(* Q: 고르기 → 응답 필터 → 제한 (지령원 Q 제한 + 정격 + 제한 모듈 Q). 다른 경로 몫을 합쳐 제한 (Auto만) *)
stQRng := F_RangeOpen();
IF _stApply.bSrcLimit THEN
	stQRng := _stQSrcLim;		// 지령원 Q 제한 (P와 같음: Manual은 정책 bSrcLimit). 접속점 기준 → 설비 기준 (보정만큼 옮김)
	IF stQRng.nMaxModule <> 0 THEN stQRng.fMax := stQRng.fMax + fQComp; END_IF
	IF stQRng.nMinModule <> 0 THEN stQRng.fMin := stQRng.fMin + fQComp; END_IF
END_IF
IF _stApply.bRating THEN
	stQRng := F_RangeAnd(stQRng, _stEnv.stQ);
END_IF
FOR i := 1 TO GVL_PARAM.LIMIT_COUNT DO
	// Q도 P와 같은 규칙: 설비 기준 모듈은 bDevLimit, 접속점 기준 모듈은 M_PccLimitOn (Manual은 bPccLimit + 모듈 bManual)
	// Q 범위는 설비 기준(접속점 + 보정)이므로 접속점 기준 모듈 값은 보정만큼 옮겨 겹침 (P는 보정 앞 단계에서 자름)
	IF M_DevLimitOn(i) THEN
		stQRng := F_RangeAdd(stQRng, _astLim[i].stQ, _anLimModule[i]);
	ELSIF M_PccLimitOn(i) THEN
		stQLim		:= _astLim[i].stQ;
		stQLim.fMax	:= stQLim.fMax + fQComp;
		stQLim.fMin	:= stQLim.fMin + fQComp;
		stQRng := F_RangeAdd(stQRng, stQLim, _anLimModule[i]);
	END_IF
END_FOR
stDiag.stQRng		:= stQRng;
stDiag.bQGroupCmd	:= _stGrpQ.bActive;
stDiag.bQUnitCmd	:= _bUnitQCmd;
tTau := T#0S;
IF _stApply.bRamp THEN
	tTau := _tQFilter;
END_IF
// 목표 = 그룹 지령 (필터 후 + 보정). 없으면 유닛 지령 합 + 다른 경로 몫 (필터는 그 값을 따라가게만 둠)
IF _stGrpQ.bActive THEN
	_afbQFilter[i_nGroup](i_fIn := _stGrpQ.fValue, i_tTau := tTau);
	stDiag.stQ := F_RangeClamp(_afbQFilter[i_nGroup].q_fOut + fQComp, stQRng);
ELSE
	_afbQFilter[i_nGroup](i_fIn := _fUnitQSum + _fOtherQ - fQComp, i_tTau := tTau);
	stDiag.stQ := F_RangeClamp(_fUnitQSum + _fOtherQ, stQRng);
END_IF
M_ShapePath := stDiag;
END_METHOD

METHOD PRIVATE M_PccLimitOn : BOOL		// 이번 경로에 접속점 기준 모듈 i를 적용하는가
VAR_INPUT
	i_nLimit	: UINT;
END_VAR
M_PccLimitOn := _abLimOn[i_nLimit] AND _aeBasis[i_nLimit] = E_LimitBasis.Pcc
				AND (NOT i_bManual OR (_stApply.bPccLimit AND _abPccManual[i_nLimit]));
END_METHOD

METHOD PRIVATE M_DevLimitOn : BOOL		// 이번 경로에 설비 기준 모듈 i를 적용하는가 (Manual은 정책 bDevLimit)
VAR_INPUT
	i_nLimit	: UINT;
END_VAR
M_DevLimitOn := _stApply.bDevLimit AND _abLimOn[i_nLimit] AND _aeBasis[i_nLimit] = E_LimitBasis.Device;
END_METHOD

METHOD PRIVATE M_TraceSet		// 추적표에 한 줄 추가
VAR_INPUT
	i_eStep		: E_TraceStep;
	i_fValue	: REAL;
	i_nModule	: UINT;
	i_bCut		: BOOL;
END_VAR
IF _stTrace.nCount < GVL_PARAM.TRACE_STEP_MAX - 2 THEN		// 끝 두 줄(분배 후·쓴 값)은 FB_OutputDiag 몫
	_stTrace.nCount := _stTrace.nCount + 1;
	_stTrace.astStep[_stTrace.nCount].eStep		:= i_eStep;
	_stTrace.astStep[_stTrace.nCount].fValue	:= i_fValue;
	_stTrace.astStep[_stTrace.nCount].bCut		:= i_bCut;
	_stTrace.astStep[_stTrace.nCount].nModule	:= i_nModule;
	_stTrace.astStep[_stTrace.nCount].nReason	:= 0;
END_IF
END_METHOD

METHOD PRIVATE M_TraceClamp : REAL		// 범위 하나로 자르고 추적표에 한 줄. 자른 값을 돌려줌
VAR_INPUT
	i_eStep		: E_TraceStep;
	i_fIn		: REAL;
	i_stRange	: ST_Range;
END_VAR
VAR
	stClamp		: ST_Clamp;
END_VAR
stClamp := F_RangeClamp(i_fIn, i_stRange);
M_TraceSet(i_eStep, stClamp.fOut, stClamp.nModule, stClamp.bClamped);
IF _stTrace.nCount >= 1 THEN
	_stTrace.astStep[_stTrace.nCount].nReason := stClamp.nReason;
END_IF
M_TraceClamp := stClamp.fOut;
END_METHOD

END_FUNCTION_BLOCK

// ---- 10_Core/02_Util/FB_Lpf.TcPOU
FUNCTION_BLOCK FB_Lpf		// 1차 지연 필터
VAR_INPUT
	i_fIn			: REAL;
	i_tTau			: TIME;		// 시정수. T#0S면 필터 없이 통과
	i_bSync			: BOOL;		// 내부 값을 i_fSyncValue로 맞춤
	i_fSyncValue	: REAL;
END_VAR
VAR_OUTPUT
	q_fOut			: REAL;
END_VAR
VAR
	_fState			: REAL;
END_VAR
VAR_TEMP
	fDt				: REAL;		// s
	fTau			: REAL;		// s
END_VAR

fDt		:= F_CycleSec();
fTau	:= TIME_TO_REAL(i_tTau) / 1000.0;

IF i_bSync THEN
	_fState := i_fSyncValue;
ELSIF fTau <= 0 THEN
	_fState := i_fIn;
ELSE
	_fState := _fState + (fDt / (fTau + fDt)) * (i_fIn - _fState);
END_IF

q_fOut := _fState;

END_FUNCTION_BLOCK

// ---- 10_Core/02_Util/F_CycleSec.TcPOU
FUNCTION F_CycleSec : REAL		// 지금 태스크의 주기 (s)
VAR
	nTask		: DINT;
END_VAR

nTask := GETCURTASKINDEXEX();
F_CycleSec := UDINT_TO_REAL(TwinCAT_SystemInfoVarList._TaskInfo[nTask].CycleTime) * 1.0E-7;	// 100 ns 단위

END_FUNCTION

// ---- 10_Core/02_Util/F_RampStep.TcPOU
FUNCTION F_RampStep : REAL		// 기준값에서 한 스캔 동안 갈 수 있는 만큼만 목표 쪽으로
VAR_INPUT
	i_fTarget	: REAL;
	i_fRef		: REAL;			// 기준 (지난 스캔 최종 출력)
	i_fUpRate	: REAL;			// |값|이 커지는 쪽 (단위/s). 0 = 램프 없음
	i_fDnRate	: REAL;			// |값|이 작아지는 쪽 (단위/s). 0 = 램프 없음
END_VAR
VAR
	fRate		: REAL;
	fStep		: REAL;
END_VAR

IF ABS(i_fTarget) > ABS(i_fRef) AND i_fTarget * i_fRef >= 0 THEN
	fRate := i_fUpRate;
ELSE
	fRate := i_fDnRate;
END_IF

IF fRate <= 0 THEN
	F_RampStep := i_fTarget;
ELSE
	fStep		:= fRate * F_CycleSec();
	F_RampStep	:= i_fRef + LIMIT(-fStep, i_fTarget - i_fRef, fStep);
END_IF

END_FUNCTION

// ---- 10_Core/40_Arbitration/F_RangeClamp.TcPOU
FUNCTION F_RangeClamp : ST_Clamp		// 값을 범위 안으로. 상·하한이 겹치면 상한이 이김
VAR_INPUT
	i_fIn		: REAL;
	i_stRange	: ST_Range;
END_VAR

F_RangeClamp.fIn	:= i_fIn;
F_RangeClamp.fOut	:= i_fIn;
IF F_RangeClamp.fOut < i_stRange.fMin THEN
	F_RangeClamp.fOut		:= i_stRange.fMin;
	F_RangeClamp.bClamped	:= TRUE;
	F_RangeClamp.nModule	:= i_stRange.nMinModule;
	F_RangeClamp.nReason	:= i_stRange.nMinReason;
END_IF
IF F_RangeClamp.fOut > i_stRange.fMax THEN
	F_RangeClamp.fOut		:= i_stRange.fMax;
	F_RangeClamp.bClamped	:= TRUE;
	F_RangeClamp.nModule	:= i_stRange.nMaxModule;
	F_RangeClamp.nReason	:= i_stRange.nMaxReason;
END_IF

END_FUNCTION

// ---- 10_Core/50_Distribution/FB_Distributor.TcPOU
FUNCTION_BLOCK FB_Distributor		// 유닛에 나눔: 경로마다(Manual → Auto) 유닛 지령 → 그룹 몫 → 유닛 지령 축소, 그다음 배터리 그룹(방향·순 한도) → 피상전력
// Auto·Manual이 같은 순서 (M_DistPath). 그룹 지령이 없으면 그룹 몫은 0 (지령 없는 유닛은 0). 유닛 지령은 성형 결과(제한)에 걸릴 때만 줄임
// Manual 정책에서 정격·BMS 한도를 끈 Manual 유닛은 그 한도를 안 씀 (bRating을 끄면 유닛 제한 모듈만 씀)
// 유닛·버스 한도는 FB_EquipmentLimits 결과. 버스 한도는 나누는 동안 남은 한도로 보고(넘친 몫은 다른 유닛에 재분배), 끝에 한 번 더 확인
// 그룹 몫을 나누는 무게는 분배 정책(그룹마다 I_DistPolicy, 비우면 코어 기본 FB_DistStd = eDistBasis). 음수·이상값 무게는 0
VAR_IN_OUT
	iq_aipDistPolicy	: ARRAY[1..GVL_PARAM.GROUP_COUNT] OF I_DistPolicy;	// 그룹별 분배 정책 (GVL_SITE.g_aipDistPolicy)
END_VAR
VAR_IN_OUT CONSTANT
	(* Auto 경로 (fbAutoShape·fbAutoGate) *)
	iq_afAutoGrpP		: ARRAY[1..GVL_PARAM.GROUP_COUNT] OF REAL;
	iq_afAutoGrpQ		: ARRAY[1..GVL_PARAM.GROUP_COUNT] OF REAL;
	iq_afAutoUnitP		: ARRAY[1..GVL_PARAM.UNIT_COUNT] OF REAL;
	iq_afAutoUnitQ		: ARRAY[1..GVL_PARAM.UNIT_COUNT] OF REAL;
	iq_astAutoUnitP		: ARRAY[1..GVL_PARAM.UNIT_COUNT] OF ST_Pick;		// 유닛별 값이 있는지
	iq_astAutoUnitQ		: ARRAY[1..GVL_PARAM.UNIT_COUNT] OF ST_Pick;
	iq_abAutoGrpPCmd	: ARRAY[1..GVL_PARAM.GROUP_COUNT] OF BOOL;		// Auto 그룹 P 지령 있음 (fbAutoShape.q_abGrpPCmd)
	iq_abAutoGrpQCmd	: ARRAY[1..GVL_PARAM.GROUP_COUNT] OF BOOL;
	(* Manual 경로 (fbManualShape·fbManualGate) *)
	iq_afManualGrpP		: ARRAY[1..GVL_PARAM.GROUP_COUNT] OF REAL;
	iq_afManualGrpQ		: ARRAY[1..GVL_PARAM.GROUP_COUNT] OF REAL;
	iq_afManualUnitP	: ARRAY[1..GVL_PARAM.UNIT_COUNT] OF REAL;
	iq_afManualUnitQ	: ARRAY[1..GVL_PARAM.UNIT_COUNT] OF REAL;
	iq_astManualUnitP	: ARRAY[1..GVL_PARAM.UNIT_COUNT] OF ST_Pick;
	iq_astManualUnitQ	: ARRAY[1..GVL_PARAM.UNIT_COUNT] OF ST_Pick;
	iq_abManualGrpPCmd	: ARRAY[1..GVL_PARAM.GROUP_COUNT] OF BOOL;		// Manual 그룹 P 지령 있음 (fbManualShape.q_abGrpPCmd)
	iq_abManualGrpQCmd	: ARRAY[1..GVL_PARAM.GROUP_COUNT] OF BOOL;
	iq_astManualPolicy	: ARRAY[1..GVL_PARAM.GROUP_COUNT] OF ST_ManualPolicy;
	(* 공통 *)
	iq_abOutputReady	: ARRAY[1..GVL_PARAM.UNIT_COUNT] OF BOOL;	// 유닛 출력 가능 = 분배 대상 (FB_OutputReady)
	iq_aeNotReadyBy	: ARRAY[1..GVL_PARAM.UNIT_COUNT] OF E_UnitLimitBy;	// 못 내는 이유
	iq_aeOpMode		: ARRAY[1..GVL_PARAM.UNIT_COUNT] OF E_OpMode;
	iq_astUnitEnv	: ARRAY[1..GVL_PARAM.UNIT_COUNT] OF ST_UnitEnvelope;	// 유닛 한도 (FB_EquipmentLimits)
	iq_astBatEnv	: ARRAY[1..GVL_PARAM.BAT_COUNT] OF ST_BatEnvelope;	// 버스 한도 (FB_EquipmentLimits)
	iq_astUnitCfg	: ARRAY[1..GVL_PARAM.UNIT_COUNT] OF ST_UnitCfg;
	iq_astBatGroup	: ARRAY[1..GVL_PARAM.BAT_COUNT] OF ST_BatGroupState;
	iq_astGroupSet	: ARRAY[1..GVL_PARAM.GROUP_COUNT] OF ST_GroupSet;
END_VAR
VAR_OUTPUT
	q_astUnitSet	: ARRAY[1..GVL_PARAM.UNIT_COUNT] OF ST_PQ;		// 유닛 최종 지령
	q_astUnitDiag	: ARRAY[1..GVL_PARAM.UNIT_COUNT] OF ST_UnitDiag;
	q_astDistDiag	: ARRAY[1..GVL_PARAM.GROUP_COUNT] OF ST_DistDiag;
	q_astBatDiag	: ARRAY[1..GVL_PARAM.BAT_COUNT] OF ST_BatDistDiag;
	q_abUnitLimited	: ARRAY[1..GVL_PARAM.UNIT_COUNT] OF BOOL;		// 유닛 지령이 요청보다 줄었거나 0으로 묶임 (P 또는 Q). 제어용: Manual 재전송 판단 (FB_Dispatcher)
	q_abManualLimitOff: ARRAY[1..GVL_PARAM.GROUP_COUNT] OF BOOL;		// Manual 정책에서 정격·BMS 한도 중 하나라도 꺼짐 (HMI 표시용)
END_VAR
VAR
	(* 유닛 사본·작업값 (메서드에서 씀) *)
	_anGroup		: ARRAY[1..GVL_PARAM.UNIT_COUNT] OF UINT;
	_anBat			: ARRAY[1..GVL_PARAM.UNIT_COUNT] OF UINT;
	_abInDist		: ARRAY[1..GVL_PARAM.UNIT_COUNT] OF BOOL;		// 출력 가능 (FB_OutputReady)
	_abManual		: ARRAY[1..GVL_PARAM.UNIT_COUNT] OF BOOL;
	_abPFix			: ARRAY[1..GVL_PARAM.UNIT_COUNT] OF BOOL;		// 자기 경로에 유닛별 P 값 있음
	_abQFix			: ARRAY[1..GVL_PARAM.UNIT_COUNT] OF BOOL;
	_afPUnitReq		: ARRAY[1..GVL_PARAM.UNIT_COUNT] OF REAL;		// 자기 경로 유닛별 값 (성형 후)
	_afQUnitReq		: ARRAY[1..GVL_PARAM.UNIT_COUNT] OF REAL;
	_abNoRating		: ARRAY[1..GVL_PARAM.UNIT_COUNT] OF BOOL;		// Manual 정책: 정격·Derate·피상전력 안 씀
	_abNoBatLimit	: ARRAY[1..GVL_PARAM.UNIT_COUNT] OF BOOL;		// Manual 정책: BMS 충방전 한도 안 씀
	_astUnitEnv	: ARRAY[1..GVL_PARAM.UNIT_COUNT] OF ST_UnitEnvelope;	// 유닛 한도 사본 (메서드에서 씀)
	_astBatEnv	: ARRAY[1..GVL_PARAM.BAT_COUNT] OF ST_BatEnvelope;	// 버스 한도 사본
	_afBusDisLeft	: ARRAY[1..GVL_PARAM.BAT_COUNT] OF REAL;	// 버스 방전 쪽 남은 한도 (양수, 나누는 동안 줄어듦. 여러 그룹이 같은 버스를 써도 한 번만 씀)
	_afBusChgLeft	: ARRAY[1..GVL_PARAM.BAT_COUNT] OF REAL;	// 버스 충전 쪽 남은 한도 (양수)
	_anPModule	: ARRAY[1..GVL_PARAM.UNIT_COUNT] OF UINT;	// P를 줄인 모듈 (유닛 제한·버스 제한 모듈. 0 = 코어)
	_afPMax			: ARRAY[1..GVL_PARAM.UNIT_COUNT] OF REAL;
	_afPMin			: ARRAY[1..GVL_PARAM.UNIT_COUNT] OF REAL;
	_afQMax			: ARRAY[1..GVL_PARAM.UNIT_COUNT] OF REAL;
	_afQMin			: ARRAY[1..GVL_PARAM.UNIT_COUNT] OF REAL;
	_afPRated		: ARRAY[1..GVL_PARAM.UNIT_COUNT] OF REAL;
	_afQRated		: ARRAY[1..GVL_PARAM.UNIT_COUNT] OF REAL;
	_afSoc			: ARRAY[1..GVL_PARAM.UNIT_COUNT] OF REAL;		// 연결 배터리 그룹 SOC (%). 모르면 -1
	_afPWork		: ARRAY[1..GVL_PARAM.UNIT_COUNT] OF REAL;
	_afQWork		: ARRAY[1..GVL_PARAM.UNIT_COUNT] OF REAL;
	_aePBy			: ARRAY[1..GVL_PARAM.UNIT_COUNT] OF E_UnitLimitBy;
	_aeQBy			: ARRAY[1..GVL_PARAM.UNIT_COUNT] OF E_UnitLimitBy;
	_afPWeight		: ARRAY[1..GVL_PARAM.UNIT_COUNT] OF REAL;		// P 몫을 나눌 때 쓴 무게 (진단)
	_abBatNoChg		: ARRAY[1..GVL_PARAM.UNIT_COUNT] OF BOOL;		// 연결 배터리 버스 충전 한도 0 → 충전 몫 안 줌
	_abBatNoDis		: ARRAY[1..GVL_PARAM.UNIT_COUNT] OF BOOL;		// 방전 한도 0 → 방전 몫 안 줌
	_eBasis			: E_DistBasis;		// 지금 그룹의 분배 기준
	_fbDistStd		: FB_DistStd;		// 코어 기본 분배 정책
	_aipDistPolicy	: ARRAY[1..GVL_PARAM.GROUP_COUNT] OF I_DistPolicy;	// 사본 (메서드에서 씀)
END_VAR
VAR_TEMP
	u				: UINT;
	g				: UINT;
	b				: UINT;
	
	fScale			: REAL;
	fBusNetP		: REAL;
	fManualNetP		: REAL;			// 버스의 Manual 유닛 P 합 (버스 방향은 Manual 우선)
	fBusDir			: REAL;			// 정한 버스 방향 (+ 방전, − 충전, 0 = 정할 수 없음)
	bHasPos			: BOOL;
	bHasNeg			: BOOL;
	fBusLimit		: REAL;
	fSLimit			: REAL;
	fFill			: REAL;			// Auto가 채울 Manual 부족분 (Auto 그룹 지령이 있을 때만)
	stDist			: ST_DistDiag;
	stBat			: ST_BatDistDiag;
END_VAR

_aipDistPolicy := iq_aipDistPolicy;
(* 0) 유닛 준비: 운전 대상, 자기 경로 값, 유닛 한도 (FB_EquipmentLimits) *)
FOR u := 1 TO GVL_PARAM.UNIT_COUNT DO
	_anGroup[u]		:= iq_astUnitCfg[u].nGroup;
	_anBat[u]		:= iq_astUnitCfg[u].nBatGroup;
	g				:= _anGroup[u];
	// 분배 대상 = 출력 가능 유닛 (FB_OutputReady. 못 내는 유닛에 몫을 주지 않음)
	_abInDist[u]	:= iq_abOutputReady[u];
	_abManual[u]	:= iq_aeOpMode[u] = E_OpMode.Manual;
	IF _abManual[u] THEN
		_abPFix[u]		:= iq_astManualUnitP[u].bActive;
		_abQFix[u]		:= iq_astManualUnitQ[u].bActive;
		_afPUnitReq[u]	:= iq_afManualUnitP[u];
		_afQUnitReq[u]	:= iq_afManualUnitQ[u];
	ELSE
		_abPFix[u]		:= iq_astAutoUnitP[u].bActive;
		_abQFix[u]		:= iq_astAutoUnitQ[u].bActive;
		_afPUnitReq[u]	:= iq_afAutoUnitP[u];
		_afQUnitReq[u]	:= iq_afAutoUnitQ[u];
	END_IF
	_abNoRating[u]		:= FALSE;
	_abNoBatLimit[u]	:= FALSE;
	IF _abManual[u] AND g >= 1 AND g <= GVL_PARAM.GROUP_COUNT THEN
		_abNoRating[u]		:= NOT iq_astManualPolicy[g].bRating;
		_abNoBatLimit[u]	:= NOT iq_astManualPolicy[g].bBatLimit;
	END_IF
	_astUnitEnv[u]	:= iq_astUnitEnv[u];
	_afPRated[u]	:= iq_astUnitCfg[u].fPRated;
	_afQRated[u]	:= iq_astUnitCfg[u].fQRated;
	// 유닛 한도 = 정격 × Derate ∩ 유닛 제한 모듈. Manual 정책 bRating을 끈 유닛은 유닛 제한 모듈만
	IF NOT _abInDist[u] THEN
		_afPMax[u]	:= 0;
		_afPMin[u]	:= 0;
		_afQMax[u]	:= 0;
		_afQMin[u]	:= 0;
	ELSIF _abNoRating[u] THEN
		_afPMax[u]	:= MIN(_astUnitEnv[u].stPRule.fMax, GVL_CORE.NO_LIMIT);
		_afPMin[u]	:= MAX(_astUnitEnv[u].stPRule.fMin, -GVL_CORE.NO_LIMIT);
		_afQMax[u]	:= MIN(_astUnitEnv[u].stQRule.fMax, GVL_CORE.NO_LIMIT);
		_afQMin[u]	:= MAX(_astUnitEnv[u].stQRule.fMin, -GVL_CORE.NO_LIMIT);
	ELSE
		_afPMax[u]	:= _astUnitEnv[u].stP.fMax;
		_afPMin[u]	:= _astUnitEnv[u].stP.fMin;
		_afQMax[u]	:= _astUnitEnv[u].stQ.fMax;
		_afQMin[u]	:= _astUnitEnv[u].stQ.fMin;
	END_IF

	_afSoc[u] := -1;
	_abBatNoChg[u] := FALSE;
	_abBatNoDis[u] := FALSE;
	b := _anBat[u];
	IF b >= 1 AND b <= GVL_PARAM.BAT_COUNT THEN
		IF iq_astBatGroup[b].stSoc.bValid THEN
			_afSoc[u] := iq_astBatGroup[b].stSoc.fValue;
		END_IF
		// 배터리 버스가 그 방향을 못 받으면 유닛 한도를 미리 0 → 나눌 때 다른 유닛으로 넘어감
		IF NOT _abNoBatLimit[u] THEN
			_abBatNoChg[u] := iq_astBatEnv[b].stP.fMin >= 0;
			_abBatNoDis[u] := iq_astBatEnv[b].stP.fMax <= 0;
		END_IF
		IF _abBatNoChg[u] THEN
			_afPMin[u] := 0;
		END_IF
		IF _abBatNoDis[u] THEN
			_afPMax[u] := 0;
		END_IF
	END_IF

	_afPWork[u] := 0;
	_afQWork[u] := 0;
	_afPWeight[u] := 0;
	_anPModule[u] := 0;
	_aePBy[u] := iq_aeNotReadyBy[u];	// 출력 못 내는 이유 (FB_OutputReady)
	_aeQBy[u] := _aePBy[u];
END_FOR

(* 버스 남은 한도: 나누는 동안 유닛에 준 만큼 줄어듦 (방전·충전 쪽 따로. 여러 그룹이 같은 버스를 써도 한 번만 씀) *)
FOR b := 1 TO GVL_PARAM.BAT_COUNT DO
	_astBatEnv[b]	:= iq_astBatEnv[b];
	_afBusDisLeft[b]	:= MAX(iq_astBatEnv[b].stP.fMax, 0.0);
	_afBusChgLeft[b]	:= MAX(-iq_astBatEnv[b].stP.fMin, 0.0);
END_FOR
(* 1) 제어 그룹마다 나누기: Manual 경로 먼저, Auto 경로는 Manual이 덜 나간 만큼 더해서 *)
FOR g := 1 TO GVL_PARAM.GROUP_COUNT DO
	_eBasis := iq_astGroupSet[g].eDistBasis;
	q_abManualLimitOff[g] := NOT (iq_astManualPolicy[g].bRating AND iq_astManualPolicy[g].bBatLimit);

	stDist.stManualP	:= M_DistPath(g, TRUE, FALSE, iq_afManualGrpP[g], iq_abManualGrpPCmd[g]);
	// Manual이 덜 나간 만큼 Auto가 채우는 것은 Auto 그룹 지령(접속점 기준)이 있을 때만. 유닛 지령만 있으면 Auto 유닛 지령을 그대로 둠
	fFill := 0;
	IF iq_abAutoGrpPCmd[g] THEN
		fFill := iq_afManualGrpP[g] - stDist.stManualP.fOut;
	END_IF
	stDist.stAutoP		:= M_DistPath(g, FALSE, FALSE, iq_afAutoGrpP[g] + fFill, iq_abAutoGrpPCmd[g]);
	stDist.stManualQ	:= M_DistPath(g, TRUE, TRUE, iq_afManualGrpQ[g], iq_abManualGrpQCmd[g]);
	fFill := 0;
	IF iq_abAutoGrpQCmd[g] THEN
		fFill := iq_afManualGrpQ[g] - stDist.stManualQ.fOut;
	END_IF
	stDist.stAutoQ		:= M_DistPath(g, FALSE, TRUE, iq_afAutoGrpQ[g] + fFill, iq_abAutoGrpQCmd[g]);
	q_astDistDiag[g]	:= stDist;
END_FOR

FOR u := 1 TO GVL_PARAM.UNIT_COUNT DO
	q_astUnitDiag[u].fPReq := _afPWork[u];
	q_astUnitDiag[u].fQReq := _afQWork[u];
END_FOR

(* 2) 배터리 그룹(DC 버스)마다 마지막 확인: 순 방향과 반대인 유닛은 0, 그다음 순 한도 (BMS 한도를 끈 Manual 유닛은 순 한도에서 뺌)
   한도는 나누는 동안 이미 맞췄으므로 보통은 줄이지 않음 (유닛별 값이 서로 반대 방향일 때 등) *)
FOR b := 1 TO GVL_PARAM.BAT_COUNT DO
	fBusNetP	:= 0;
	fManualNetP	:= 0;
	bHasPos		:= FALSE;
	bHasNeg		:= FALSE;
	FOR u := 1 TO GVL_PARAM.UNIT_COUNT DO
		IF _anBat[u] = b THEN
			fBusNetP := fBusNetP + _afPWork[u];
			IF _abManual[u] THEN fManualNetP := fManualNetP + _afPWork[u]; END_IF
			bHasPos := bHasPos OR _afPWork[u] > 0;
			bHasNeg := bHasNeg OR _afPWork[u] < 0;
		END_IF
	END_FOR
	stBat.fNetIn	:= fBusNetP;
	stBat.nDirZero	:= 0;
	stBat.fScale	:= 1.0;
	// 버스 방향: Manual 유닛 쪽 순 방향이 먼저 (Manual 우선), 없으면 전체 순 방향. 둘 다 0이면 정할 수 없으므로 반대 방향끼리 모두 0 (버스 안 순환 방지)
	fBusDir := fManualNetP;
	IF ABS(fBusDir) <= 0.01 THEN fBusDir := fBusNetP; END_IF
	IF ABS(fBusDir) <= 0.01 THEN fBusDir := 0; END_IF
	FOR u := 1 TO GVL_PARAM.UNIT_COUNT DO
		IF _anBat[u] = b AND ((fBusDir > 0 AND _afPWork[u] < 0) OR (fBusDir < 0 AND _afPWork[u] > 0)
			OR (fBusDir = 0 AND bHasPos AND bHasNeg AND _afPWork[u] <> 0)) THEN
			_afPWork[u]		:= 0;
			_aePBy[u]		:= E_UnitLimitBy.BatDir;
			stBat.nDirZero	:= stBat.nDirZero + 1;
		END_IF
	END_FOR

	fBusNetP := 0;
	FOR u := 1 TO GVL_PARAM.UNIT_COUNT DO
		IF _anBat[u] = b AND NOT _abNoBatLimit[u] THEN fBusNetP := fBusNetP + _afPWork[u]; END_IF
	END_FOR
	IF fBusNetP > 0 THEN
		fBusLimit := iq_astBatEnv[b].stP.fMax;
	ELSE
		fBusLimit := iq_astBatEnv[b].stP.fMin;
	END_IF
	stBat.fNetDir	:= fBusNetP;
	stBat.fLimit	:= fBusLimit;
	IF (fBusNetP > 0 AND fBusNetP > fBusLimit) OR (fBusNetP < 0 AND fBusNetP < fBusLimit) THEN
		fScale := fBusLimit / fBusNetP;
		stBat.fScale := fScale;
		FOR u := 1 TO GVL_PARAM.UNIT_COUNT DO
			IF _anBat[u] = b AND NOT _abNoBatLimit[u] AND _afPWork[u] <> 0 THEN
				_afPWork[u]	:= _afPWork[u] * fScale;
				_aePBy[u]	:= E_UnitLimitBy.BatLimit;
				IF fBusNetP > 0 THEN
					_anPModule[u] := iq_astBatEnv[b].stP.nMaxModule;
				ELSE
					_anPModule[u] := iq_astBatEnv[b].stP.nMinModule;
				END_IF
			END_IF
		END_FOR
	END_IF
	q_astBatDiag[b] := stBat;
END_FOR

FOR u := 1 TO GVL_PARAM.UNIT_COUNT DO
	q_astUnitDiag[u].fPBat := _afPWork[u];
END_FOR

(* 3) 피상전력: 우선이 아닌 쪽을 줄임 (다른 유닛에 다시 나누지 않음). 정격을 끈 Manual 유닛은 건너뜀 *)
FOR u := 1 TO GVL_PARAM.UNIT_COUNT DO
	g := _anGroup[u];
	fSLimit := _astUnitEnv[u].fSMax;
	IF _abInDist[u] AND NOT _abNoRating[u] AND fSLimit > 0 AND g >= 1 AND g <= GVL_PARAM.GROUP_COUNT
		AND (_afPWork[u] * _afPWork[u] + _afQWork[u] * _afQWork[u]) > fSLimit * fSLimit THEN
		IF iq_astGroupSet[g].bQPriority THEN
			_afQWork[u]	:= LIMIT(-fSLimit, _afQWork[u], fSLimit);
			_afPWork[u]	:= SEL(_afPWork[u] < 0, 1.0, -1.0) * SQRT(MAX(0.0, fSLimit * fSLimit - _afQWork[u] * _afQWork[u]));
			_aePBy[u]	:= E_UnitLimitBy.SLimit;
		ELSE
			_afPWork[u]	:= LIMIT(-fSLimit, _afPWork[u], fSLimit);
			_afQWork[u]	:= SEL(_afQWork[u] < 0, 1.0, -1.0) * SQRT(MAX(0.0, fSLimit * fSLimit - _afPWork[u] * _afPWork[u]));
			_aeQBy[u]	:= E_UnitLimitBy.SLimit;
		END_IF
	END_IF
END_FOR

(* 4) 출력 *)
FOR u := 1 TO GVL_PARAM.UNIT_COUNT DO
	q_astUnitSet[u].fP			:= _afPWork[u];
	q_astUnitSet[u].fQ			:= _afQWork[u];
	IF _abPFix[u] THEN
		q_astUnitDiag[u].eRole	:= E_UnitRole.Fixed;
	ELSIF _abManual[u] THEN
		q_astUnitDiag[u].eRole	:= E_UnitRole.ManualShare;
	ELSE
		q_astUnitDiag[u].eRole	:= E_UnitRole.AutoShare;
	END_IF
	q_astUnitDiag[u].fPOut		:= _afPWork[u];
	q_astUnitDiag[u].ePBy	:= _aePBy[u];
	q_astUnitDiag[u].nPModule	:= _anPModule[u];
	q_astUnitDiag[u].fQOut		:= _afQWork[u];
	q_astUnitDiag[u].eQBy		:= _aeQBy[u];
	q_astUnitDiag[u].fPMax		:= _afPMax[u];
	q_astUnitDiag[u].fPWeight	:= _afPWeight[u];
	q_abUnitLimited[u]			:= M_IsLimited(_aePBy[u]) OR M_IsLimited(_aeQBy[u]);
END_FOR

METHOD PRIVATE M_DistPath : ST_DistPathDiag		// 경로 하나(Auto 또는 Manual)의 P 또는 Q를 나눔. 두 경로가 같은 순서
// ① 유닛별 값 (유닛 한도) → ② 그룹 지령이 있으면 남은 양을 그룹 몫 유닛에 (그룹 목표와 반대 방향으로는 안 감) → ③ 그래도 넘치면 유닛별 값을 비율로 줄임 (늘리지는 않음)
VAR_INPUT
	i_nGroup	: UINT;
	i_bManual	: BOOL;
	i_bForQ		: BOOL;
	i_fTarget	: REAL;			// 이 경로 목표 (성형 결과)
	i_bGrpCmd	: BOOL;			// 이 경로 그룹 지령 있음
END_VAR
VAR
	u			: UINT;
	bFix		: BOOL;
	fFixed		: REAL;
	fShareReq	: REAL;
	fShareGot	: REAL;
	fScale		: REAL;
	fOut		: REAL;
	stDiag		: ST_DistPathDiag;
	(* [결함 5 수정 2026-11-03: 추가] 유닛별 P 값을 버스마다 같은 비율로 줄이는 데 씀 *)
	b			: UINT;
	fVal		: REAL;
	afFixP		: ARRAY[1..GVL_PARAM.UNIT_COUNT] OF REAL;	// 유닛 한도 안으로 넣은 유닛별 P
	afFixDis	: ARRAY[1..GVL_PARAM.BAT_COUNT] OF REAL;	// 버스별 유닛별 P 합 (방전 쪽, 양수)
	afFixChg	: ARRAY[1..GVL_PARAM.BAT_COUNT] OF REAL;	// 버스별 유닛별 P 합 (충전 쪽, 양수)
	afScDis		: ARRAY[1..GVL_PARAM.BAT_COUNT] OF REAL;	// 버스별 비율 (방전 쪽, 1 = 안 줄임)
	afScChg		: ARRAY[1..GVL_PARAM.BAT_COUNT] OF REAL;
END_VAR
// ① 유닛별 값
fFixed := 0;
// [결함 5 수정 2026-11-03: P 유닛별 값은 버스마다 합을 먼저 보고, 남은 버스 한도를 넘으면 그 버스 유닛 값을 같은 비율로 줄임 (이유 BatLimit).
//   원래는 유닛 순서로 M_SetP(u, M_ClampToBus(u, M_ClampToUnitLimit(u, FALSE, _afPUnitReq[u]))) → 앞 유닛이 남은 한도를 다 씀]
FOR b := 1 TO GVL_PARAM.BAT_COUNT DO
	afFixDis[b]	:= 0;
	afFixChg[b]	:= 0;
	afScDis[b]	:= 1.0;
	afScChg[b]	:= 1.0;
END_FOR
FOR u := 1 TO GVL_PARAM.UNIT_COUNT DO
	bFix := SEL(i_bForQ, _abPFix[u], _abQFix[u]);
	IF _anGroup[u] = i_nGroup AND _abInDist[u] AND _abManual[u] = i_bManual AND bFix THEN
		IF i_bForQ THEN
			_afQWork[u]	:= M_ClampToUnitLimit(u, TRUE, _afQUnitReq[u]);
			fFixed		:= fFixed + _afQWork[u];
		ELSE
			afFixP[u]	:= M_ClampToUnitLimit(u, FALSE, _afPUnitReq[u]);
			b			:= _anBat[u];
			IF b >= 1 AND b <= GVL_PARAM.BAT_COUNT AND NOT _abNoBatLimit[u] THEN
				afFixDis[b]	:= afFixDis[b] + MAX(afFixP[u], 0.0);
				afFixChg[b]	:= afFixChg[b] + MAX(-afFixP[u], 0.0);
			END_IF
		END_IF
	END_IF
END_FOR
IF NOT i_bForQ THEN
	FOR b := 1 TO GVL_PARAM.BAT_COUNT DO
		IF afFixDis[b] > MAX(_afBusDisLeft[b], 0.0) + 0.01 THEN afScDis[b] := MAX(_afBusDisLeft[b], 0.0) / afFixDis[b]; END_IF
		IF afFixChg[b] > MAX(_afBusChgLeft[b], 0.0) + 0.01 THEN afScChg[b] := MAX(_afBusChgLeft[b], 0.0) / afFixChg[b]; END_IF
	END_FOR
	FOR u := 1 TO GVL_PARAM.UNIT_COUNT DO
		IF _anGroup[u] = i_nGroup AND _abInDist[u] AND _abManual[u] = i_bManual AND _abPFix[u] THEN
			fVal	:= afFixP[u];
			b		:= _anBat[u];
			IF b >= 1 AND b <= GVL_PARAM.BAT_COUNT AND NOT _abNoBatLimit[u] THEN
				IF fVal > 0 AND afScDis[b] < 1.0 THEN
					fVal := fVal * afScDis[b];
					M_MarkBusLimit(u, TRUE);
				ELSIF fVal < 0 AND afScChg[b] < 1.0 THEN
					fVal := fVal * afScChg[b];
					M_MarkBusLimit(u, FALSE);
				END_IF
			END_IF
			M_SetP(u, M_ClampToBus(u, fVal));
			fFixed	:= fFixed + _afPWork[u];
		END_IF
	END_FOR
END_IF

// ② 그룹 몫
fShareReq := i_fTarget - fFixed;
IF NOT i_bGrpCmd THEN
	fShareReq := 0.0;						// 그룹 지령 없음: 지령 없는 유닛에는 안 줌
ELSIF i_fTarget >= 0 THEN
	fShareReq := MAX(fShareReq, 0.0);
ELSE
	fShareReq := MIN(fShareReq, 0.0);
END_IF
fShareGot := M_SplitToShareUnits(i_nGroup, i_bManual, i_bForQ, fShareReq);

// ③ 유닛별 값 축소
fScale := 1.0;
IF fFixed <> 0 THEN
	fScale := LIMIT(0.0, (i_fTarget - fShareGot) / fFixed, 1.0);
END_IF
IF fScale < 1.0 THEN
	FOR u := 1 TO GVL_PARAM.UNIT_COUNT DO
		bFix := SEL(i_bForQ, _abPFix[u], _abQFix[u]);
		IF _anGroup[u] = i_nGroup AND _abInDist[u] AND _abManual[u] = i_bManual AND bFix THEN
			IF i_bForQ THEN
				_afQWork[u]	:= _afQWork[u] * fScale;
				_aeQBy[u]	:= E_UnitLimitBy.Scaled;
			ELSE
				M_SetP(u, _afPWork[u] * fScale);
				_aePBy[u]	:= E_UnitLimitBy.Scaled;
			END_IF
		END_IF
	END_FOR
END_IF

fOut := 0;
FOR u := 1 TO GVL_PARAM.UNIT_COUNT DO
	IF _anGroup[u] = i_nGroup AND _abManual[u] = i_bManual THEN
		fOut := fOut + SEL(i_bForQ, _afPWork[u], _afQWork[u]);
	END_IF
END_FOR

stDiag.fTarget		:= i_fTarget;
stDiag.fFixed		:= fFixed;
stDiag.fShareReq	:= fShareReq;
stDiag.fShareGot	:= fShareGot;
stDiag.fFixedScale	:= fScale;
stDiag.fOut			:= fOut;
M_DistPath := stDiag;
END_METHOD

METHOD PRIVATE M_IsLimited : BOOL		// 이 이유가 "요청보다 줄었거나 0으로 묶임"인가 (이유를 추가하면 여기서 정함. 열거 순서에 기대지 않음)
VAR_INPUT
	i_eBy		: E_UnitLimitBy;
END_VAR
CASE i_eBy OF
	E_UnitLimitBy.Rating, E_UnitLimitBy.Derate, E_UnitLimitBy.Scaled, E_UnitLimitBy.BatDir, E_UnitLimitBy.BatLimit,
	E_UnitLimitBy.SLimit, E_UnitLimitBy.ModeSwitch, E_UnitLimitBy.WaitManualCmd, E_UnitLimitBy.UnitRule:
		M_IsLimited := TRUE;
ELSE
	M_IsLimited := FALSE;		// None, NotAvail, NotRun (출력 없음은 Run 들어감·나옴으로 따로 씀)
END_CASE
END_METHOD

METHOD PRIVATE M_ClampToUnitLimit : REAL	// 유닛 한도(설비 한도) 안으로
VAR_INPUT
	i_nUnit		: UINT;
	i_bForQ		: BOOL;
	i_fValue		: REAL;
END_VAR
VAR
	fUnitMax		: REAL;
	fUnitMin		: REAL;
END_VAR
IF i_bForQ THEN
	fUnitMax := _afQMax[i_nUnit];
	fUnitMin := _afQMin[i_nUnit];
ELSE
	fUnitMax := _afPMax[i_nUnit];
	fUnitMin := _afPMin[i_nUnit];
END_IF

M_ClampToUnitLimit := LIMIT(fUnitMin, i_fValue, fUnitMax);
IF M_ClampToUnitLimit <> i_fValue THEN
	M_MarkUnitLimitReason(i_nUnit, i_bForQ, i_fValue);
END_IF
END_METHOD

METHOD PRIVATE M_MarkUnitLimitReason	// 유닛 한도에 걸린 이유 기록 (어느 쪽 한도를 무엇이 정했나)
VAR_INPUT
	i_nUnit	: UINT;
	i_bForQ	: BOOL;
	i_fDir	: REAL;	// 요청 방향 (+ 방전·공급, - 충전·흡수)
END_VAR
VAR
	eLimitBy	: E_UnitLimitBy;
	stRng	: ST_Range;
END_VAR
IF NOT i_bForQ AND ((i_fDir < 0 AND _abBatNoChg[i_nUnit]) OR (i_fDir > 0 AND _abBatNoDis[i_nUnit])) THEN
	M_MarkBusLimit(i_nUnit, i_fDir > 0);
	RETURN;
END_IF
IF i_bForQ THEN
	IF _abNoRating[i_nUnit] THEN
		stRng := _astUnitEnv[i_nUnit].stQRule;
	ELSE
		stRng := _astUnitEnv[i_nUnit].stQ;
	END_IF
	IF i_fDir > 0 THEN eLimitBy := _astUnitEnv[i_nUnit].eQMaxBy; ELSE eLimitBy := _astUnitEnv[i_nUnit].eQMinBy; END_IF
ELSE
	IF _abNoRating[i_nUnit] THEN
		stRng := _astUnitEnv[i_nUnit].stPRule;
	ELSE
		stRng := _astUnitEnv[i_nUnit].stP;
	END_IF
	IF i_fDir > 0 THEN eLimitBy := _astUnitEnv[i_nUnit].ePMaxBy; ELSE eLimitBy := _astUnitEnv[i_nUnit].ePMinBy; END_IF
END_IF
IF _abNoRating[i_nUnit] THEN
	eLimitBy := E_UnitLimitBy.UnitRule;		// 정격을 안 쓰는 유닛은 유닛 제한 모듈에만 걸림
END_IF
IF i_bForQ THEN
	_aeQBy[i_nUnit] := eLimitBy;
ELSE
	_aePBy[i_nUnit] := eLimitBy;
	IF i_fDir > 0 THEN
		_anPModule[i_nUnit] := stRng.nMaxModule;
	ELSE
		_anPModule[i_nUnit] := stRng.nMinModule;
	END_IF
END_IF
END_METHOD

METHOD PRIVATE M_ShareWeight : REAL		// 분배 무게: 그룹 분배 정책 (없으면 코어 기본). 음수·이상값은 0
VAR_INPUT
	i_nUnit		: UINT;
	i_bForQ		: BOOL;
	i_bPositive	: BOOL;			// 나눌 양이 방전·공급 쪽
END_VAR
VAR
	stView	: ST_DistView;
	g		: UINT;
	fW		: REAL;
END_VAR
g := _anGroup[i_nUnit];
stView.nGroup		:= g;
stView.nUnit		:= i_nUnit;
stView.bManual		:= _abManual[i_nUnit];
stView.bForQ		:= i_bForQ;
stView.bPositive	:= i_bPositive;
stView.eBasis		:= _eBasis;
stView.fPRated		:= _afPRated[i_nUnit];
stView.fQRated		:= _afQRated[i_nUnit];
stView.fSoc			:= _afSoc[i_nUnit];
IF g >= 1 AND g <= GVL_PARAM.GROUP_COUNT AND_THEN _aipDistPolicy[g] <> 0 THEN
	fW := _aipDistPolicy[g].M_Weight(i_stView := stView);
ELSE
	fW := _fbDistStd.M_Weight(i_stView := stView);
END_IF
// NaN·무한대를 먼저 거름 (OR는 단락 평가가 아니라서 fW < 0을 NaN으로 비교하지 않게 나눔)
IF NOT F_CmdOk(fW, 0.0) THEN
	fW := 0.0;
ELSIF fW < 0.0 THEN
	fW := 0.0;
END_IF
M_ShareWeight := fW;
END_METHOD

METHOD PRIVATE M_SplitToShareUnits : REAL	// 그룹 몫 유닛에 무게대로 나눔. 한도에 걸린 유닛 몫은 나머지에 다시. 실제로 나눈 양을 돌려줌
// P는 연결 버스 남은 한도도 봄: 한 라운드에 한 버스로 가는 몫이 남은 한도보다 크면 그 버스 유닛 몫을 같은 비율로 줄이고(공평하게), 그 유닛들은 다 찬 것으로 뺌 → 넘친 몫은 다른 버스 유닛에
VAR_INPUT
	i_nGroup	: UINT;
	i_bManual	: BOOL;			// TRUE = Manual 그룹 몫 유닛, FALSE = Auto 그룹 몫 유닛
	i_bForQ		: BOOL;
	i_fAmount	: REAL;
END_VAR
VAR
	u			: UINT;
	nRound		: UINT;
	bPositive		: BOOL;
	fRemaining		: REAL;
	fWeightSum		: REAL;
	fAssigned		: REAL;
	fNewValue		: REAL;
	fUnitCap		: REAL;
	abCanTake	: ARRAY[1..GVL_PARAM.UNIT_COUNT] OF BOOL;
	bBusCap	: BOOL;	// 이번 상한이 버스 남은 한도 때문
	b	: UINT;
	fBusScale	: REAL;	// 이 유닛 몫에 곱하는 버스 비율 (1 = 안 줄임)
	afBusWant	: ARRAY[1..GVL_PARAM.BAT_COUNT] OF REAL;	// 이번 라운드 버스별 요청 증가량 (양수)
	afBusScale	: ARRAY[1..GVL_PARAM.BAT_COUNT] OF REAL;	// 버스별 비율
	bCut		: BOOL;	// 한도 때문에 이번 몫보다 덜 받음. [결함 5 수정 2026-11-03: 추가]
	bBusScaled	: BOOL;	// 이번 라운드 버스 비율로 줄었음. [결함 5 수정 2026-11-03: 추가]
END_VAR
bPositive := i_fAmount >= 0;

// 대상 유닛: 이 그룹, 운전 대상, 같은 운전 모드, 그 값(P 또는 Q)에 유닛별 값이 없는 유닛
FOR u := 1 TO GVL_PARAM.UNIT_COUNT DO
	abCanTake[u] := _anGroup[u] = i_nGroup AND _abInDist[u] AND (_abManual[u] = i_bManual)
				AND ((i_bForQ AND NOT _abQFix[u]) OR (NOT i_bForQ AND NOT _abPFix[u]));
END_FOR

fRemaining := i_fAmount;
FOR nRound := 1 TO GVL_PARAM.UNIT_COUNT DO
	IF ABS(fRemaining) < 0.001 THEN
		EXIT;
	END_IF
	fWeightSum := 0;
	FOR u := 1 TO GVL_PARAM.UNIT_COUNT DO
		IF abCanTake[u] THEN fWeightSum := fWeightSum + M_ShareWeight(u, i_bForQ, bPositive); END_IF
	END_FOR
	IF fWeightSum <= 0 THEN
		EXIT;	// 더 받을 유닛이 없음
	END_IF
	// P: 버스별 요청 증가량이 남은 한도보다 크면 그 버스 몫을 비율로 줄임
	FOR b := 1 TO GVL_PARAM.BAT_COUNT DO
		afBusWant[b]	:= 0;
		afBusScale[b]	:= 1.0;
	END_FOR
	IF NOT i_bForQ THEN
		FOR u := 1 TO GVL_PARAM.UNIT_COUNT DO
			b := _anBat[u];
			IF abCanTake[u] AND b >= 1 AND b <= GVL_PARAM.BAT_COUNT AND NOT _abNoBatLimit[u] THEN
				afBusWant[b] := afBusWant[b] + ABS(fRemaining) * M_ShareWeight(u, FALSE, bPositive) / fWeightSum;
			END_IF
		END_FOR
		FOR b := 1 TO GVL_PARAM.BAT_COUNT DO
			IF bPositive AND afBusWant[b] > _afBusDisLeft[b] THEN
				afBusScale[b] := MAX(_afBusDisLeft[b], 0.0) / afBusWant[b];
			ELSIF NOT bPositive AND afBusWant[b] > _afBusChgLeft[b] THEN
				afBusScale[b] := MAX(_afBusChgLeft[b], 0.0) / afBusWant[b];
			END_IF
		END_FOR
	END_IF

	fAssigned := 0;
	FOR u := 1 TO GVL_PARAM.UNIT_COUNT DO
		IF abCanTake[u] THEN
			IF i_bForQ THEN
				fNewValue := _afQWork[u] + fRemaining * M_ShareWeight(u, i_bForQ, bPositive) / fWeightSum;
				fUnitCap := SEL(bPositive, _afQMin[u], _afQMax[u]);
				bBusCap := FALSE;
				fBusScale := 1.0;
			ELSE
				_afPWeight[u] := M_ShareWeight(u, i_bForQ, bPositive);
				fBusScale := 1.0;
				b := _anBat[u];
				IF b >= 1 AND b <= GVL_PARAM.BAT_COUNT AND NOT _abNoBatLimit[u] THEN
					fBusScale := afBusScale[b];
				END_IF
				fNewValue := _afPWork[u] + fRemaining * _afPWeight[u] / fWeightSum * fBusScale;
				// 유닛 한도와 연결 버스 남은 한도 중 좁은 쪽
				fUnitCap := SEL(bPositive, MAX(_afPMin[u], M_BusMin(u)), MIN(_afPMax[u], M_BusMax(u)));
				bBusCap := fUnitCap <> SEL(bPositive, _afPMin[u], _afPMax[u]);
			END_IF
			IF (bPositive AND fNewValue >= fUnitCap) OR (NOT bPositive AND fNewValue <= fUnitCap) THEN
				// [결함 5 수정 2026-11-03: 이유는 실제로 덜 받았을 때만 (몫이 한도를 넘었거나 버스 비율로 줄었을 때). 몫이 한도에 딱 닿기만 하면 안 남김.
				//   원래 IF ABS(fRemaining) > 0.001 THEN (버스 한도 ELSE 유닛 한도) → 같은 몫인데 마지막 유닛만 BatLimit로 나옴]
				bCut			:= ABS(fNewValue - fUnitCap) > 0.01;
				bBusScaled		:= NOT i_bForQ AND fBusScale < 0.9999;
				fNewValue		:= fUnitCap;
				abCanTake[u]	:= FALSE;
				IF bCut AND NOT bBusCap THEN
					M_MarkUnitLimitReason(u, i_bForQ, SEL(bPositive, -1.0, 1.0));
				ELSIF bCut OR bBusScaled THEN
					M_MarkBusLimit(u, bPositive);
				END_IF
			END_IF
			IF i_bForQ THEN
				fAssigned	:= fAssigned + fNewValue - _afQWork[u];
				_afQWork[u]	:= fNewValue;
			ELSE
				fAssigned	:= fAssigned + fNewValue - _afPWork[u];
				M_SetP(u, fNewValue);
			END_IF
		END_IF
	END_FOR
	fRemaining := fRemaining - fAssigned;
	// 남은 한도를 다 쓴 버스의 유닛만 뺌. 버스 비율로 줄였어도 한도가 남으면(같은 버스 다른 유닛이 자기 한도에 먼저 걸림) 다음 라운드에 더 받음
	IF NOT i_bForQ THEN
		FOR u := 1 TO GVL_PARAM.UNIT_COUNT DO
			b := _anBat[u];
			IF abCanTake[u] AND b >= 1 AND b <= GVL_PARAM.BAT_COUNT AND NOT _abNoBatLimit[u]
				AND ((bPositive AND _afBusDisLeft[b] <= 0.001) OR (NOT bPositive AND _afBusChgLeft[b] <= 0.001)) THEN
				abCanTake[u] := FALSE;
				IF ABS(fRemaining) > 0.001 THEN
					M_MarkBusLimit(u, bPositive);
				END_IF
			END_IF
		END_FOR
	END_IF
END_FOR

M_SplitToShareUnits := i_fAmount - fRemaining;
END_METHOD

METHOD PRIVATE M_SetP	// 유닛 P를 바꾸고 연결 버스 남은 한도를 맞춤 (방전·충전 쪽 따로)
VAR_INPUT
	i_nUnit	: UINT;
	i_fNew	: REAL;
END_VAR
VAR
	b	: UINT;
	fOld	: REAL;
END_VAR
fOld := _afPWork[i_nUnit];
b := _anBat[i_nUnit];
IF b >= 1 AND b <= GVL_PARAM.BAT_COUNT AND NOT _abNoBatLimit[i_nUnit] THEN
	_afBusDisLeft[b] := _afBusDisLeft[b] + MAX(fOld, 0.0) - MAX(i_fNew, 0.0);
	_afBusChgLeft[b] := _afBusChgLeft[b] + MAX(-fOld, 0.0) - MAX(-i_fNew, 0.0);
END_IF
_afPWork[i_nUnit] := i_fNew;
END_METHOD

METHOD PRIVATE M_BusMax : REAL	// 이 유닛이 가질 수 있는 P 상한 (연결 버스 남은 방전 한도 기준). 버스 한도를 안 보는 유닛은 아주 큰 값
VAR_INPUT
	i_nUnit	: UINT;
END_VAR
VAR
	b	: UINT;
END_VAR
b := _anBat[i_nUnit];
IF b >= 1 AND b <= GVL_PARAM.BAT_COUNT AND NOT _abNoBatLimit[i_nUnit] THEN
	M_BusMax := MAX(_afPWork[i_nUnit], 0.0) + MAX(_afBusDisLeft[b], 0.0);
ELSE
	M_BusMax := GVL_CORE.NO_LIMIT;
END_IF
END_METHOD

METHOD PRIVATE M_BusMin : REAL	// 이 유닛이 가질 수 있는 P 하한 (연결 버스 남은 충전 한도 기준)
VAR_INPUT
	i_nUnit	: UINT;
END_VAR
VAR
	b	: UINT;
END_VAR
b := _anBat[i_nUnit];
IF b >= 1 AND b <= GVL_PARAM.BAT_COUNT AND NOT _abNoBatLimit[i_nUnit] THEN
	M_BusMin := MIN(_afPWork[i_nUnit], 0.0) - MAX(_afBusChgLeft[b], 0.0);
ELSE
	M_BusMin := -GVL_CORE.NO_LIMIT;
END_IF
END_METHOD

METHOD PRIVATE M_ClampToBus : REAL	// 유닛별 P를 연결 버스 남은 한도 안으로 (값은 M_SetP로 씀)
VAR_INPUT
	i_nUnit	: UINT;
	i_fValue	: REAL;
END_VAR
M_ClampToBus := LIMIT(M_BusMin(i_nUnit), i_fValue, M_BusMax(i_nUnit));
IF M_ClampToBus <> i_fValue THEN
	M_MarkBusLimit(i_nUnit, i_fValue > 0);
END_IF
END_METHOD

METHOD PRIVATE M_MarkBusLimit	// 버스 한도에 걸림: 이유 BatLimit, 그 쪽 한도를 정한 모듈 (0 = BMS 한도)
VAR_INPUT
	i_nUnit	: UINT;
	i_bDis	: BOOL;	// 방전 쪽
END_VAR
VAR
	b	: UINT;
END_VAR
_aePBy[i_nUnit] := E_UnitLimitBy.BatLimit;
b := _anBat[i_nUnit];
IF b >= 1 AND b <= GVL_PARAM.BAT_COUNT THEN
	IF i_bDis THEN
		_anPModule[i_nUnit] := _astBatEnv[b].stP.nMaxModule;
	ELSE
		_anPModule[i_nUnit] := _astBatEnv[b].stP.nMinModule;
	END_IF
END_IF
END_METHOD

END_FUNCTION_BLOCK

// ---- 10_Core/50_Distribution/FB_DistStd.TcPOU
FUNCTION_BLOCK FB_DistStd EXTENDS FB_ModuleBase IMPLEMENTS I_DistPolicy	// 코어 기본 분배: 그룹 설정 eDistBasis (정격 비율 / SOC / 균등)

METHOD M_Weight : REAL
VAR_INPUT
	i_stView	: ST_DistView;
END_VAR
IF i_stView.eBasis = E_DistBasis.Equal THEN
	M_Weight := 1.0;
ELSIF i_stView.eBasis = E_DistBasis.Soc AND NOT i_stView.bForQ AND i_stView.fSoc >= 0 THEN
	IF i_stView.bPositive THEN
		M_Weight := MAX(i_stView.fSoc, 1.0);			// 방전: SOC 높은 쪽
	ELSE
		M_Weight := MAX(100.0 - i_stView.fSoc, 1.0);	// 충전: SOC 낮은 쪽
	END_IF
ELSIF i_stView.bForQ THEN
	M_Weight := i_stView.fQRated;
ELSE
	M_Weight := i_stView.fPRated;
END_IF
END_METHOD

END_FUNCTION_BLOCK

// ---- 10_Core/60_Dispatch/FB_Sequencer.TcPOU
FUNCTION_BLOCK FB_Sequencer		// 유닛·BMS 시퀀서를 묶음: 이번 스캔 조건, 접수 검사, 유닛·BMS 명령 (배터리 요청 정리는 FB_BatRequest, 기동 조건은 FB_PermitEval, 그룹 상태는 FB_GroupState)
// 호출 순서 (MAIN): M_Prepare(이번 스캔 조건) → M_CheckRequest(접수 검사) → 본체(분배 뒤, 실제 단계 진행·명령 생성)
VAR_INPUT
	i_bTestReset	: BOOL;			// 시험: 모든 PCS·BMS 고장 리셋 (TEST_MODE에서만 MAIN이 넘김)
	i_bCmdEnable	: BOOL := TRUE;	// FALSE = 설정 오류: 명령을 만들지 않음
	i_bWriteEnable	: BOOL := TRUE;	// FALSE = 장비 쓰기 불가 (DEVICE_WRITE 꺼짐·대기 PLC): 명령을 만들지 않고 기동 요청은 WriteDisabled로 거부
END_VAR
VAR_IN_OUT CONSTANT
	iq_abNewReq		: ARRAY[1..GVL_PARAM.UNIT_COUNT] OF BOOL;		// 이번 스캔에 접수된 지령원 상태 요청 있음 (FB_StateArbiter)
	iq_aeReq		: ARRAY[1..GVL_PARAM.UNIT_COUNT] OF E_PcsCmd;	// 그 요청
	iq_astUnitProt	: ARRAY[1..GVL_PARAM.UNIT_COUNT] OF ST_UnitProt;	// 보호 결과: 정지·비상정지는 시퀀서가 보냄 (보호 명령만 재시도)
	iq_aeStartMode	: ARRAY[1..GVL_PARAM.UNIT_COUNT] OF E_StartMode;
	iq_astUnit		: ARRAY[1..GVL_PARAM.UNIT_COUNT] OF ST_UnitState;
	iq_astAvail		: ARRAY[1..GVL_PARAM.UNIT_COUNT] OF ST_UnitAvail;
	iq_astUnitCfg	: ARRAY[1..GVL_PARAM.UNIT_COUNT] OF ST_UnitCfg;
	iq_astBms		: ARRAY[1..GVL_PARAM.BMS_COUNT] OF ST_BatState;
	iq_astBmsCfg	: ARRAY[1..GVL_PARAM.BMS_COUNT] OF ST_BmsCfg;
	iq_astBmsAvail	: ARRAY[1..GVL_PARAM.BMS_COUNT] OF ST_BmsAvail;
	iq_astBmsProt	: ARRAY[1..GVL_PARAM.BMS_COUNT] OF ST_BmsProt;
	iq_astSrcOut	: ARRAY[1..GVL_PARAM.SOURCE_COUNT] OF ST_SourceOutput;	// 지령원 배터리 요청 (FB_BatRequest로), 고장 리셋 요청
	iq_astReg		: ARRAY[1..GVL_PARAM.SOURCE_COUNT] OF ST_SourceReg;
	iq_aeOpMode		: ARRAY[1..GVL_PARAM.UNIT_COUNT] OF E_OpMode;			// 실제 운전 모드
	iq_stSet		: ST_SeqSet;
END_VAR
VAR_OUTPUT
	q_astUnitCmd	: ARRAY[1..GVL_PARAM.UNIT_COUNT] OF ST_PcsCmd;
	q_astBmsCmd		: ARRAY[1..GVL_PARAM.BMS_COUNT] OF ST_BatCmd;
	q_abWaitPermit	: ARRAY[1..GVL_PARAM.GROUP_COUNT] OF BOOL;		// 그룹에 기동 조건을 기다리는 유닛 있음 (FB_PermitEval이 다음 스캔에 씀)
	(* 진단 *)
	q_aeUnitSeq		: ARRAY[1..GVL_PARAM.UNIT_COUNT] OF E_UnitSeq;
	q_abAccept		: ARRAY[1..GVL_PARAM.UNIT_COUNT] OF BOOL;		// 접수 검사 결과: 이번 스캔 후보를 받음 (FB_StateArbiter.M_CommitRequest로)
	q_aeRefuse		: ARRAY[1..GVL_PARAM.UNIT_COUNT] OF E_SeqRefuse;	// 마지막 기동 쪽 요청 거부 이유 (받아들이면 None)
	q_abStopping	: ARRAY[1..GVL_PARAM.UNIT_COUNT] OF BOOL;		// 정지 진행 중 (출력 0. FB_OutputReady가 다음 스캔에 씀)
	q_aeFailCmd		: ARRAY[1..GVL_PARAM.UNIT_COUNT] OF E_PcsCmd;	// 확인되지 않은 명령 (실패 알람, 잠그지 않음)
	q_aeBatRefuse	: ARRAY[1..GVL_PARAM.BAT_COUNT] OF E_SeqRefuse;		// 배터리 그룹별 마지막 요청 거부 이유 (FB_BatRequest)
	q_abBatHoldOpen	: ARRAY[1..GVL_PARAM.BAT_COUNT] OF BOOL;		// 지령원 BatOpen으로 연 배터리 그룹 (FB_BatRequest)
	q_abBatRefusedNow: ARRAY[1..GVL_PARAM.BAT_COUNT] OF BOOL;		// 이번 스캔에 배터리 요청을 거부함 (1스캔, 로그용)
	q_abBatReqTaken	: ARRAY[1..GVL_PARAM.SOURCE_COUNT] OF BOOL;		// 지령원의 이번 배터리 요청을 받은 배터리 그룹이 있음 (로그용)
	q_aeBmsFailCmd	: ARRAY[1..GVL_PARAM.BMS_COUNT] OF E_BatCmd;	// 확인되지 않은 BMS 명령 (실패 알람, 잠그지 않음)
END_VAR
VAR
	_afbUnit		: ARRAY[1..GVL_PARAM.UNIT_COUNT] OF FB_UnitSeq;
	_afbBms			: ARRAY[1..GVL_PARAM.BMS_COUNT] OF FB_BmsSeq;
	_fbBatReq		: FB_BatRequest;
	(* 이번 스캔 조건 (M_Prepare). 접수 검사와 본체가 같은 값을 씀 *)
	_bCtxCmdEnable	: BOOL;
	_bCtxWriteEnable: BOOL;
	_abCtxComm		: ARRAY[1..GVL_PARAM.UNIT_COUNT] OF BOOL;
	_aeCtxRun		: ARRAY[1..GVL_PARAM.UNIT_COUNT] OF E_RunState;
	_abCtxAvail		: ARRAY[1..GVL_PARAM.UNIT_COUNT] OF BOOL;
	_abCtxBatReady	: ARRAY[1..GVL_PARAM.UNIT_COUNT] OF BOOL;		// 연결 배터리 그룹 투입 완료 (배터리 없는 유닛은 TRUE)
	_abCtxPermit	: ARRAY[1..GVL_PARAM.UNIT_COUNT] OF BOOL;		// 그룹 기동 조건
	_aeCtxStartMode	: ARRAY[1..GVL_PARAM.UNIT_COUNT] OF E_StartMode;
	_abCtxInstalled	: ARRAY[1..GVL_PARAM.UNIT_COUNT] OF BOOL;		// 유닛 설치됨 (PCS 칸 있음). [결함 6 수정 2026-11-03: 추가]
END_VAR
VAR_TEMP
	u				: UINT;
	m				: UINT;
	g				: UINT;
	b				: UINT;
	abWantBat		: ARRAY[1..GVL_PARAM.BAT_COUNT] OF BOOL;
	eProtCmd		: E_PcsCmd;
	i				: UINT;
	bUnitReset		: BOOL;
	abBatReset		: ARRAY[1..GVL_PARAM.BAT_COUNT] OF BOOL;
END_VAR

(* 1) 이번 스캔 조건은 M_Prepare가 준비함 (MAIN이 접수 검사 전에 부름) *)
FOR g := 1 TO GVL_PARAM.GROUP_COUNT DO
	q_abWaitPermit[g] := FALSE;
END_FOR

(* 2) 유닛 시퀀서 *)
// 고장 리셋은 장비에 내리는 명령일 뿐: 지령원 PCS Reset(대상 유닛, 0 = 대상 그룹 전체) → 그 PCS, 배터리 Reset(대상 배터리 그룹, 0 = 전체) → 그 그룹 BMS
FOR b := 1 TO GVL_PARAM.BAT_COUNT DO
	abWantBat[b]	:= FALSE;
	abBatReset[b]	:= i_bTestReset;
	FOR i := 1 TO GVL_PARAM.SOURCE_COUNT DO
		IF iq_astSrcOut[i].bValid AND iq_astSrcOut[i].stBatReq.eCmd = E_BatCmd.Reset
			AND (iq_astSrcOut[i].stBatReq.nBatGroup = 0 OR iq_astSrcOut[i].stBatReq.nBatGroup = b) THEN
			abBatReset[b] := TRUE;
		END_IF
	END_FOR
END_FOR
FOR u := 1 TO GVL_PARAM.UNIT_COUNT DO
	g := iq_astUnitCfg[u].nGroup;
	b := iq_astUnitCfg[u].nBatGroup;

	bUnitReset := i_bTestReset;
	FOR i := 1 TO GVL_PARAM.SOURCE_COUNT DO
		IF iq_astSrcOut[i].bValid AND iq_astSrcOut[i].stPcsReq.eCmd = E_PcsCmd.Reset
			AND (iq_astReg[i].nGroup = 0 OR iq_astReg[i].nGroup = g)
			AND (iq_astSrcOut[i].stPcsReq.nUnit = 0 OR iq_astSrcOut[i].stPcsReq.nUnit = u) THEN
			bUnitReset := TRUE;
		END_IF
	END_FOR
	// 보호 정지 쪽 조치만 명령으로 (보호 대기 = 출력 0, 가용 아님으로 이미 빠짐)
	CASE iq_astUnitProt[u].ePcsAction OF
		E_PcsAction.Stop:	eProtCmd := E_PcsCmd.Stop;
		E_PcsAction.EStop:	eProtCmd := E_PcsCmd.EStop;
	ELSE
		eProtCmd := E_PcsCmd.None;
	END_CASE
	_afbUnit[u](i_bNewReq		:= iq_abNewReq[u],
				i_eReq			:= iq_aeReq[u],
				i_eProtCmd		:= eProtCmd,
				i_bProtActive	:= iq_astUnitProt[u].ePcsAction <> E_PcsAction.None,
				i_eStartMode	:= iq_aeStartMode[u],
				i_stUnit		:= iq_astUnit[u],
				i_bAvail		:= iq_astAvail[u].bAvail,
				i_bBatReady		:= _abCtxBatReady[u],
				i_bPermit		:= _abCtxPermit[u],
				i_fPRated		:= iq_astUnitCfg[u].fPRated,
				i_bReset		:= bUnitReset,
				i_bCmdEnable	:= i_bCmdEnable AND i_bWriteEnable,
				i_stSet			:= iq_stSet.stPcs);
	q_astUnitCmd[u]		:= _afbUnit[u].q_stCmd;
	q_aeUnitSeq[u]		:= _afbUnit[u].q_eSeqState;
	q_aeFailCmd[u]		:= _afbUnit[u].q_eFailCmd;
	q_abStopping[u]		:= _afbUnit[u].q_bStopping;

	IF b >= 1 AND b <= GVL_PARAM.BAT_COUNT AND _afbUnit[u].q_bWantBat AND iq_stSet.stBat.eClose <> E_BatClose.OnRequest THEN
		abWantBat[b] := TRUE;
	END_IF
	IF g >= 1 AND g <= GVL_PARAM.GROUP_COUNT AND _afbUnit[u].q_bWaitPermit THEN
		q_abWaitPermit[g] := TRUE;
	END_IF
END_FOR

(* 3) 배터리 요청 정리 (지령원 BatClose·BatOpen, 정지 시 개방, 운전원이 연 배터리 유지) *)
_fbBatReq(	i_bOpenOnStop	:= iq_stSet.stBat.bOpenOnStop,
			iq_astSrcOut	:= iq_astSrcOut,
			iq_astReg		:= iq_astReg,
			iq_aeOpMode		:= iq_aeOpMode,
			iq_astUnitCfg	:= iq_astUnitCfg,
			iq_astUnit		:= iq_astUnit,
			iq_abNewReq		:= iq_abNewReq,
			iq_aeReq		:= iq_aeReq,
			iq_abWantBat	:= abWantBat);
q_aeBatRefuse		:= _fbBatReq.q_aeRefuse;
q_abBatHoldOpen		:= _fbBatReq.q_abHoldOpen;
q_abBatRefusedNow	:= _fbBatReq.q_abRefusedNow;
q_abBatReqTaken		:= _fbBatReq.q_abReqTaken;

(* 4) BMS 시퀀서 *)
FOR m := 1 TO GVL_PARAM.BMS_COUNT DO
	b := iq_astBmsCfg[m].nBatGroup;
	IF b >= 1 AND b <= GVL_PARAM.BAT_COUNT THEN
		_afbBms[m](	i_bWantClose	:= abWantBat[b] AND NOT _fbBatReq.q_abHoldOpen[b],
					i_bCloseReq		:= _fbBatReq.q_abCloseReq[b],
					i_bOpenReq		:= _fbBatReq.q_abOpenReq[b],
					i_eProtAction	:= iq_astBmsProt[m].eBatAction,
					i_bUnitsStopped	:= _fbBatReq.q_abBusStopOk[b],
					i_bUsable		:= iq_astBmsAvail[m].bUsable,
					i_stBms			:= iq_astBms[m],
					i_bReset		:= abBatReset[b],
					i_bCmdEnable	:= i_bCmdEnable AND i_bWriteEnable,
					i_stSet			:= iq_stSet.stBat);
	END_IF
	q_astBmsCmd[m]		:= _afbBms[m].q_stCmd;
	q_aeBmsFailCmd[m]	:= _afbBms[m].q_eFailCmd;
END_FOR

METHOD M_Prepare		// 이번 스캔 조건을 한 번만 모음: 유닛 상태, 배터리 투입 완료(FB_BatGroup), 그룹 기동 조건(FB_PermitEval). 접수 검사와 본체가 같이 씀
VAR_INPUT
	i_bCmdEnable	: BOOL;
	i_bWriteEnable	: BOOL := TRUE;
END_VAR
VAR_IN_OUT CONSTANT
	iq_aeStartMode	: ARRAY[1..GVL_PARAM.UNIT_COUNT] OF E_StartMode;
	iq_astUnit		: ARRAY[1..GVL_PARAM.UNIT_COUNT] OF ST_UnitState;
	iq_astAvail		: ARRAY[1..GVL_PARAM.UNIT_COUNT] OF ST_UnitAvail;
	iq_astUnitCfg	: ARRAY[1..GVL_PARAM.UNIT_COUNT] OF ST_UnitCfg;
	iq_astBatGroup	: ARRAY[1..GVL_PARAM.BAT_COUNT] OF ST_BatGroupState;	// 투입 완료 bReady (FB_BatGroup)
	iq_abPermit		: ARRAY[1..GVL_PARAM.GROUP_COUNT] OF BOOL;				// 그룹 기동 조건 (FB_PermitEval)
	iq_abUnitInstalled	: ARRAY[1..GVL_PARAM.UNIT_COUNT] OF BOOL;			// 유닛 설치됨 (FB_ModuleList). 미설치 유닛은 요청을 안 받음 (정지에 머물고 그룹 상태에 안 걸림). [결함 6 수정 2026-11-03: 추가]
END_VAR
VAR
	u				: UINT;
	g				: UINT;
	b				: UINT;
END_VAR
FOR u := 1 TO GVL_PARAM.UNIT_COUNT DO
	g := iq_astUnitCfg[u].nGroup;
	b := iq_astUnitCfg[u].nBatGroup;
	_abCtxBatReady[u] := TRUE;							// 배터리 없는 유닛
	IF b >= 1 AND b <= GVL_PARAM.BAT_COUNT THEN
		_abCtxBatReady[u] := iq_astBatGroup[b].bReady;
	ELSIF b > GVL_PARAM.BAT_COUNT THEN
		_abCtxBatReady[u] := FALSE;						// 설정 오류
	END_IF
	_abCtxPermit[u] := TRUE;
	IF g >= 1 AND g <= GVL_PARAM.GROUP_COUNT THEN
		_abCtxPermit[u] := iq_abPermit[g];
	END_IF
	_abCtxComm[u]		:= iq_astUnit[u].bComm;
	_aeCtxRun[u]		:= iq_astUnit[u].eRunState;
	_abCtxAvail[u]		:= iq_astAvail[u].bAvail;
	_aeCtxStartMode[u]	:= iq_aeStartMode[u];
	_abCtxInstalled[u]	:= iq_abUnitInstalled[u];	// [결함 6 수정 2026-11-03: 추가]
END_FOR
_bCtxCmdEnable	:= i_bCmdEnable;
_bCtxWriteEnable	:= i_bWriteEnable;
END_METHOD

METHOD M_CheckRequest		// 접수 검사 (순수 판단): 정지 쪽은 항상 받음. 기동 쪽은 검사하고 거부 이유를 남김
// 타이머·재시도 횟수·명령은 건드리지 않음. M_Prepare 다음에 부름 (정지 진행 중은 지난 스캔 유닛 시퀀서 값)
VAR_IN_OUT CONSTANT
	iq_abCand		: ARRAY[1..GVL_PARAM.UNIT_COUNT] OF BOOL;		// FB_StateArbiter.q_abCand
	iq_aeCand		: ARRAY[1..GVL_PARAM.UNIT_COUNT] OF E_PcsCmd;	// FB_StateArbiter.q_aeCand
END_VAR
VAR
	u				: UINT;
	eRun			: E_RunState;
	bStartSide		: BOOL;
	eRefuse			: E_SeqRefuse;
END_VAR
FOR u := 1 TO GVL_PARAM.UNIT_COUNT DO
	q_abAccept[u] := FALSE;
	// [결함 6 수정 2026-11-03: 미설치 유닛은 정지 쪽도 받지 않음 (받으면 ToStop에 머물러 그룹 상태가 Stopping으로 남음). 거부 이유도 남기지 않음 (원래 IF iq_abCand[u] THEN)]
	IF iq_abCand[u] AND NOT _abCtxInstalled[u] THEN
		q_aeRefuse[u] := E_SeqRefuse.None;
	ELSIF iq_abCand[u] THEN
		eRun := _aeCtxRun[u];
		// 기동 쪽: Run, 또는 정지 상태(Stop·Fault)에서 Standby. 운전 중 Standby·Stop·EStop은 정지 쪽
		bStartSide := iq_aeCand[u] = E_PcsCmd.Run
			OR (iq_aeCand[u] = E_PcsCmd.Standby AND _abCtxComm[u] AND F_IsStopped(eRun));

		IF NOT bStartSide THEN
			q_abAccept[u] := TRUE;			// 정지 쪽은 항상 받음 (보호·코어 요청 포함)
		ELSE
			eRefuse := E_SeqRefuse.None;
			IF NOT _bCtxCmdEnable THEN
				eRefuse := E_SeqRefuse.ConfigError;
			ELSIF NOT _bCtxWriteEnable THEN
				eRefuse := E_SeqRefuse.WriteDisabled;
			ELSIF NOT _abCtxComm[u] THEN
				eRefuse := E_SeqRefuse.CommLost;
			ELSIF _afbUnit[u].q_bStopping THEN
				eRefuse := E_SeqRefuse.StopInProgress;		// 정지는 끝까지 함. 끝난 뒤 새 요청 필요
			ELSIF NOT _abCtxAvail[u] THEN
				eRefuse := E_SeqRefuse.NotAvail;
			ELSIF _aeCtxStartMode[u] <> E_StartMode.Sequence THEN
				// 단계별: 지금 단계에서 바로 할 수 있어야 함
				// 정지 → 대기(활성) 또는 Run: 배터리 투입이 먼저, Run은 기동 조건도. 이미 활성이면 할 일 없음
				IF F_IsStopped(eRun) AND NOT _abCtxBatReady[u] THEN
					eRefuse := E_SeqRefuse.NoBattery;
				ELSIF iq_aeCand[u] = E_PcsCmd.Run AND F_IsStopped(eRun) AND NOT _abCtxPermit[u] THEN
					eRefuse := E_SeqRefuse.NoPermit;
				END_IF
			END_IF
			// 순서 기동: 배터리 투입·기동 조건은 기다리는 단계라 거부하지 않음
			q_abAccept[u]		:= eRefuse = E_SeqRefuse.None;
			q_aeRefuse[u]		:= eRefuse;
		END_IF
	END_IF
END_FOR
END_METHOD

END_FUNCTION_BLOCK

// ---- 10_Core/60_Dispatch/FB_UnitSeq.TcPOU
FUNCTION_BLOCK FB_UnitSeq		// 유닛 하나의 시퀀스: 받은 명령을 한 번 보내고 장비 상태로 확인. 보호 정지 쪽 명령만 재시도
// 정지 쪽: 지령원 Stop·EStop(접수된 스캔), 보호 Stop·EStop(걸려 있는 동안) 중 센 쪽 하나. 통신이 없으면 기다렸다가 돌아오면 보냄
// 기동 쪽: 멈춘 유닛에 Run(또는 Standby = 활성 + 출력 0) 요청이 오면 Run 1회. 순서 기동은 배터리 투입 → 기동 조건 → Run
//          활성(Run·대기)이면 지령(P·Q)만 씀. PMS가 Run을 다시 보내거나 대기 명령을 만들지 않음 (대기 = 출력 0)
// 재시도: 보호 명령만 tStopRetry × nStopRetry. 넘거나 지령원 명령이 확인되지 않으면 실패 알람만 남김 (잠그지 않음)
VAR_INPUT
	i_bNewReq		: BOOL;			// 이번 스캔에 접수된 지령원 상태 요청 있음 (FB_StateArbiter)
	i_eReq			: E_PcsCmd;		// 그 요청
	i_eProtCmd		: E_PcsCmd;		// 보호 정지 쪽 조치 (Stop·EStop, 없으면 None). 보호 대기는 출력 0이라 명령 없음
	i_bProtActive	: BOOL;			// 보호 조치가 걸려 있음 (대기 포함): 진행 중인 기동을 멈춤
	i_eStartMode	: E_StartMode;
	i_stUnit		: ST_UnitState;
	i_bAvail		: BOOL;
	i_bBatReady		: BOOL;			// 연결 배터리 그룹 투입 완료 (배터리 없는 유닛은 TRUE)
	i_bPermit		: BOOL;			// 그룹 기동 조건 (등록 없으면 TRUE)
	i_fPRated		: REAL;
	i_bReset		: BOOL;			// 고장 리셋: 상승 에지에 장비가 고장이면 고장 리셋 명령 1회 (PMS 상태는 바꾸지 않음)
	i_stSet			: ST_PcsSeqSet;
	i_bCmdEnable	: BOOL := TRUE;	// FALSE = 설정 오류: 명령을 만들지 않음
END_VAR
VAR_OUTPUT
	q_stCmd			: ST_PcsCmd;		// 보낼 명령. nSeq가 바뀌면 새 명령 (디스패처가 1회 전송)
	q_eSeqState		: E_UnitSeq;
	q_bWantBat		: BOOL;			// 배터리 투입 필요 (순서 기동 중)
	q_bWaitPermit	: BOOL;			// 기동 조건 대기 중
	q_eFailCmd		: E_PcsCmd;		// 확인되지 않은 명령 (실패 알람). 새 요청이 오거나 그 보호가 풀리면 지움. None = 실패 없음
	q_bStopping		: BOOL;			// 정지 진행 중 (보낼 차례·정지 램프·확인 중). 출력 0 (FB_OutputReady), 기동 요청 거부 (접수 검사). 둘 다 다음 스캔에 씀
END_VAR
VAR
	_nCmdSeq		: UDINT;
	_ePending		: E_PcsCmd;		// 확인 중인 명령
	_bStopSide		: BOOL;			// 확인 중인 명령이 정지 쪽 (확인 시간 tStopRetry)
	_bRetry			: BOOL;			// 확인 중인 명령을 재시도함 (보호 명령)
	_nTries			: UINT;
	_eWant			: E_PcsCmd;		// 보낼 차례인 정지 쪽 명령 (통신을 기다리거나 정지 램프 중)
	_bWantRetry		: BOOL;			// 그 명령을 재시도함 (통신이 있을 때 생긴 보호 명령. 통신이 없을 때 생긴 것은 돌아오면 1회만)
	_eGaveUp		: E_PcsCmd;		// 재시도를 다 쓴 보호 명령: 그 보호가 걸려 있는 동안 다시 보내지 않음
	_bStarting		: BOOL;			// 기동 진행 중 (순서 기동은 활성이 될 때까지, 단계별은 요청 스캔만)
	_bStartPermit	: BOOL;			// 이 기동은 기동 조건을 봄 (Run 요청. Standby 요청은 안 봄)
	_tonConfirm		: TON;
	_tonStopRamp	: TON;
	_rtReset		: R_TRIG;
	_bResetReq		: BOOL;			// 고장 리셋 보낼 차례 기다림 (같은 스캔 다른 명령·진행 중인 정지가 먼저)
	(* 임시값: 본문과 액션(A_)이 함께 씀. 액션이 본문의 VAR_TEMP를 못 볼 수 있어 VAR에 둠. 매 스캔 쓴 뒤에 읽음 *)
	_eRunState		: E_RunState;
	_bRamping		: BOOL;
	_nSeqBefore		: UDINT;			// 이번 스캔 명령을 만들기 전 번호 (같은 스캔에 다른 명령을 보냈는지 확인)
END_VAR

_eRunState		:= i_stUnit.eRunState;
q_bWantBat		:= FALSE;
q_bWaitPermit	:= FALSE;
_rtReset(CLK := i_bReset);
// 실패 표시 지우기: 새 요청이 오거나, 포기한 보호 명령보다 보호가 약해지면 (다시 보낼 수 있음)
IF i_bNewReq OR F_StateRank(i_eProtCmd) < F_StateRank(_eGaveUp) THEN
	q_eFailCmd	:= E_PcsCmd.None;
	_eGaveUp	:= E_PcsCmd.None;
END_IF
IF NOT i_bCmdEnable THEN
	// 설정 오류: 명령을 만들지 않고, 진행 중인 것도 내려놓음 (기동 요청 거부는 접수 검사가 함)
	_ePending	:= E_PcsCmd.None;
	_eWant		:= E_PcsCmd.None;
	_bStarting	:= FALSE;
	_tonConfirm(IN := FALSE);
	_tonStopRamp(IN := FALSE);
	_bRamping	:= FALSE;
	_bResetReq	:= FALSE;
ELSE
	_nSeqBefore := _nCmdSeq;
	A_TakeRequest();		// 요청·보호 받기
	A_ConfirmSentCmd();		// 보낸 명령 확인
	A_SendStop();			// 정지 쪽 보내기
	A_SendStart();			// 기동 쪽 보내기
	A_ResetFault();			// 고장 리셋
END_IF
A_SummarizeState();		// 상태 요약

METHOD PRIVATE M_SendCmdAndStartConfirm	// 명령 1회 보내고 확인 시작
VAR_INPUT
	i_eCmd		: E_PcsCmd;
	i_bStopSide	: BOOL;
	i_bRetry	: BOOL;		// 확인되지 않으면 재시도 (보호 명령)
END_VAR
IF i_eCmd = _ePending THEN
	_nTries := _nTries + 1;		// 같은 명령 재전송
ELSE
	_nTries := 0;
END_IF
_nCmdSeq		:= _nCmdSeq + 1;
q_stCmd.eCmd	:= i_eCmd;
q_stCmd.nSeq	:= _nCmdSeq;
_ePending		:= i_eCmd;
_bStopSide		:= i_bStopSide;
_bRetry			:= i_bRetry;
_tonConfirm(IN := FALSE);
END_METHOD

METHOD PRIVATE M_Want	// 정지 쪽 명령을 보낼 차례로 둠: 보낼 차례인 것·확인 중인 것보다 셀 때만. 같은 명령을 확인 중이면 재시도만 더함
VAR_INPUT
	i_eCmd		: E_PcsCmd;
	i_bRetry	: BOOL;
END_VAR
IF _bStopSide AND _ePending = i_eCmd THEN
	_bRetry := _bRetry OR i_bRetry;
ELSIF F_StateRank(i_eCmd) > F_StateRank(_eWant)
	AND (NOT _bStopSide OR F_StateRank(i_eCmd) > F_StateRank(_ePending)) THEN
	_eWant		:= i_eCmd;
	_bWantRetry	:= i_bRetry;
END_IF
END_METHOD

ACTION A_TakeRequest:
(* 1) 받기: 이번 스캔에 접수된 지령원 요청, 걸려 있는 보호 *)
IF i_bNewReq THEN
	IF i_eReq = E_PcsCmd.Stop OR i_eReq = E_PcsCmd.EStop THEN
		M_Want(i_eReq, FALSE);		// 지령원 명령은 한 번만
	ELSIF (i_eReq = E_PcsCmd.Run OR i_eReq = E_PcsCmd.Standby) AND F_IsStopped(_eRunState) THEN
		// 멈춘 유닛 기동 (Standby 요청 = 활성 + 출력 0). 이미 활성이면 할 일 없음: 출력은 지령으로
		_bStarting		:= TRUE;
		_bStartPermit	:= i_eReq = E_PcsCmd.Run;
	END_IF
END_IF
// 보호 정지 쪽: 장비가 아직 그 상태가 아니면 보낼 차례로 둠. 통신이 없을 때 생긴 것은 통신이 돌아오면 1회만 (재시도 없음)
IF i_eProtCmd <> E_PcsCmd.None AND i_eProtCmd <> _eGaveUp
	AND NOT (i_stUnit.bComm AND F_CmdReached(i_eProtCmd, _eRunState)) THEN
	M_Want(i_eProtCmd, i_stUnit.bComm);
END_IF
// 보호·정지가 기동을 멈춤 (풀려도 저절로 기동하지 않음)
IF i_bProtActive OR _eWant <> E_PcsCmd.None THEN
	_bStarting := FALSE;
END_IF
END_ACTION

ACTION A_ConfirmSentCmd:
(* 2) 보낸 명령 확인: 장비 상태가 바뀌면 끝. 안 바뀌면 보호 명령만 재시도, 나머지는 실패 알람 *)
IF _ePending <> E_PcsCmd.None THEN
	IF F_CmdReached(_ePending, _eRunState) THEN
		_ePending	:= E_PcsCmd.None;
		_nTries		:= 0;
	ELSE
		IF _bStopSide THEN
			_tonConfirm(IN := TRUE, PT := i_stSet.tStopRetry);
		ELSE
			_tonConfirm(IN := TRUE, PT := i_stSet.tCmdConfirm);
		END_IF
		IF _tonConfirm.Q THEN
			IF _bRetry AND _nTries < i_stSet.nStopRetry THEN
				IF i_stUnit.bComm THEN		// 통신이 끊기면 기다렸다가 이어서 보냄 (기다린 동안은 횟수를 세지 않음)
					M_SendCmdAndStartConfirm(_ePending, _bStopSide, TRUE);
				END_IF
			ELSE
				q_eFailCmd := _ePending;		// 실패 알람만 (잠그지 않음)
				IF _bRetry THEN
					_eGaveUp := _ePending;		// 그 보호가 걸려 있는 동안 다시 보내지 않음
				END_IF
				IF NOT _bStopSide THEN
					_bStarting := FALSE;		// 기동 실패: 다시 요청해야 함
				END_IF
				_ePending := E_PcsCmd.None;
			END_IF
		END_IF
	END_IF
END_IF
END_ACTION

ACTION A_SendStop:
(* 3) 정지 쪽 보내기: 통신이 있을 때. 정지 램프를 켰으면 출력이 내려간 뒤 Stop (지령값은 q_bStopping으로 이미 0) *)
_bRamping := FALSE;
IF _eWant <> E_PcsCmd.None AND i_stUnit.bComm THEN
	IF F_CmdReached(_eWant, _eRunState) THEN
		_eWant := E_PcsCmd.None;		// 이미 그 상태
	ELSE
		IF _eWant = E_PcsCmd.Stop AND _eRunState = E_RunState.Run AND i_stSet.bStopRamp THEN
			_tonStopRamp(IN := TRUE, PT := i_stSet.tStopRampMax);
			_bRamping := ABS(i_stUnit.stP.fValue) > i_fPRated * i_stSet.fStopDonePct / 100.0 AND NOT _tonStopRamp.Q;
		END_IF
		IF NOT _bRamping THEN
			M_SendCmdAndStartConfirm(_eWant, TRUE, _bWantRetry);
			_eWant := E_PcsCmd.None;
		END_IF
	END_IF
END_IF
IF NOT _bRamping THEN
	_tonStopRamp(IN := FALSE);
END_IF
END_ACTION

ACTION A_SendStart:
(* 4) 기동 쪽: 멈춘 유닛에 Run 1회 (순서 기동은 배터리 투입 → 기동 조건 → Run). 활성(Run·대기)이 되면 끝 *)
IF _bStarting AND (_eRunState = E_RunState.Run OR _eRunState = E_RunState.Standby) THEN
	_bStarting := FALSE;
END_IF
IF _bStarting THEN
	q_bWantBat := i_eStartMode = E_StartMode.Sequence;
	IF i_bAvail AND i_stUnit.bComm AND _ePending = E_PcsCmd.None AND F_IsStopped(_eRunState) AND i_bBatReady THEN
		q_bWaitPermit := _bStartPermit AND NOT i_bPermit;
		IF NOT q_bWaitPermit THEN
			M_SendCmdAndStartConfirm(E_PcsCmd.Run, FALSE, FALSE);
		END_IF
	END_IF
	IF i_eStartMode <> E_StartMode.Sequence THEN
		_bStarting := FALSE;		// 단계별: 요청 스캔에 한 번 (배터리·기동 조건은 접수 검사가 이미 봄)
	END_IF
END_IF
END_ACTION

ACTION A_ResetFault:
(* 5) 고장 리셋: 장비가 고장이면 고장 리셋 명령 1회 (확인·재시도 없음. 풀리면 장비 상태가 Stop으로 바뀜)
   보호가 걸려 있어도 보냄. 단, 이번 스캔에 다른 명령을 보냈거나 정지가 진행 중이면 그게 끝난 뒤 보냄 (보호 명령을 덮지 않음) *)
IF _rtReset.Q THEN
	_bResetReq := TRUE;
END_IF
IF _bResetReq THEN
	IF NOT i_stUnit.bComm OR NOT (_eRunState = E_RunState.Fault OR i_stUnit.bFault) THEN
		_bResetReq := FALSE;		// 리셋할 고장 없음 (또는 통신 없음)
	ELSIF _nCmdSeq = _nSeqBefore AND NOT _bRamping AND _eWant = E_PcsCmd.None AND NOT (_ePending <> E_PcsCmd.None AND _bStopSide) THEN
		_nCmdSeq		:= _nCmdSeq + 1;
		q_stCmd.eCmd	:= E_PcsCmd.Reset;
		q_stCmd.nSeq	:= _nCmdSeq;
		_bResetReq		:= FALSE;
	END_IF
END_IF
END_ACTION

ACTION A_SummarizeState:
(* 6) 상태 요약 *)
q_bStopping := _bRamping OR _eWant <> E_PcsCmd.None OR (_ePending <> E_PcsCmd.None AND _bStopSide);
IF _bRamping THEN
	q_eSeqState := E_UnitSeq.StopRamp;
ELSIF _ePending = E_PcsCmd.Run THEN
	q_eSeqState := E_UnitSeq.ToRun;
ELSIF q_bStopping THEN
	q_eSeqState := E_UnitSeq.ToStop;
ELSIF _eRunState = E_RunState.Run THEN
	q_eSeqState := E_UnitSeq.Running;
ELSIF _eRunState = E_RunState.Standby THEN
	q_eSeqState := E_UnitSeq.Standby;
ELSIF F_IsStopped(_eRunState) THEN
	IF q_bWantBat AND NOT i_bBatReady THEN
		q_eSeqState := E_UnitSeq.WaitBat;
	ELSIF q_bWaitPermit THEN
		q_eSeqState := E_UnitSeq.WaitPermit;
	ELSE
		q_eSeqState := E_UnitSeq.Stopped;
	END_IF
ELSE
	q_eSeqState := E_UnitSeq.Unknown;
END_IF
END_ACTION

END_FUNCTION_BLOCK

// ---- 10_Core/02_Util/F_IsStopped.TcPOU
FUNCTION F_IsStopped : BOOL		// 장비가 멈춘 상태인가 (Stop 또는 Fault. Fault도 멈춘 상태). 통신 여부는 보지 않음: 통신이 있는지는 부르는 쪽이 따로 봄
VAR_INPUT
	i_eRun		: E_RunState;
END_VAR

F_IsStopped := i_eRun = E_RunState.Stop OR i_eRun = E_RunState.Fault;

END_FUNCTION

// ---- 10_Core/60_Dispatch/F_CmdReached.TcPOU
FUNCTION F_CmdReached : BOOL		// 장비 상태가 명령대로 바뀌었나
VAR_INPUT
	i_eCmd		: E_PcsCmd;
	i_eRun		: E_RunState;
END_VAR

CASE i_eCmd OF
	E_PcsCmd.Run:		F_CmdReached := i_eRun = E_RunState.Run OR i_eRun = E_RunState.Standby;	// 활성 (대기 = 활성 + 출력 0)
	E_PcsCmd.Standby:	F_CmdReached := i_eRun = E_RunState.Standby;
	E_PcsCmd.Stop,
	E_PcsCmd.EStop:	F_CmdReached := F_IsStopped(i_eRun);
ELSE
	F_CmdReached := TRUE;
END_CASE

END_FUNCTION

// ---- 10_Core/60_Dispatch/FB_BmsSeq.TcPOU
FUNCTION_BLOCK FB_BmsSeq		// BMS 하나의 접촉기: 투입은 요청·기동이 있을 때만, 개방·비상정지는 버스 유닛 정지 뒤. 보호 명령만 재시도, 실패는 알람만 (잠그지 않음)
VAR_INPUT
	i_bWantClose	: BOOL;			// 자동 투입 조건 (순서 기동 중인 유닛 있음, 투입 시점 OnStart)
	i_bCloseReq		: BOOL;			// 지령원 BatClose 요청 (이번 스캔)
	i_bOpenReq		: BOOL;			// 지령원 BatOpen 또는 정지 시 개방 (FB_BatRequest가 버스 유닛 정지를 이미 확인)
	i_eProtAction	: E_BatAction;	// 보호 조치
	i_bUnitsStopped	: BOOL;			// 같은 버스 유닛이 모두 정지 (보호 기준: Stop·Fault 보고 또는 통신 끊김)
	i_bUsable		: BOOL;			// 통신·고장·시스템 정지·보호 이상 없음
	i_stBms			: ST_BatState;
	i_bReset		: BOOL;			// 고장 리셋: 상승 에지에 BMS가 고장이면 고장 리셋 명령 1회 (PMS 상태는 바꾸지 않음)
	i_stSet			: ST_BatSeqSet;
	i_bCmdEnable	: BOOL := TRUE;	// FALSE = 설정 오류: 명령을 만들지 않음
END_VAR
VAR_OUTPUT
	q_stCmd			: ST_BatCmd;
	q_bClosed		: BOOL;
	q_eFailCmd		: E_BatCmd;		// 확인되지 않은 명령 (투입, 또는 재시도를 다 쓴 보호 개방·비상정지). 알람만. 투입 요청·새 기동·보호 변경으로 지움. None = 실패 없음
END_VAR
VAR
	_nCmdSeq		: UDINT;
	_ePending		: E_BatCmd;		// 확인 중인 명령
	_bRetry			: BOOL;			// 확인 중인 명령을 재시도함 (보호 명령)
	_nTries			: UINT;
	_tonConfirm		: TON;
	_eLastProt		: E_BatAction;
	_bProtNoComm	: BOOL;			// 보호가 걸린 동안 통신이 끊긴 적 있음: 통신이 돌아오면 1회만 보냄 (재시도 없음)
	_rtWantClose	: R_TRIG;		// 새 기동 (투입 실패 뒤 다시 투입할 수 있음)
	_rtReset		: R_TRIG;
	_bResetReq		: BOOL;			// 고장 리셋 보낼 차례 기다림 (같은 스캔 다른 명령·진행 중인 개방이 먼저)
END_VAR
VAR_TEMP
	bOpened			: BOOL;			// 개방 확인: 통신이 있고 접촉기 열림 (통신 끊김은 개방 확인 아님)
	eProtCmd		: E_BatCmd;		// 보호 조치를 명령으로
	nSeqBefore		: UDINT;
END_VAR

q_bClosed	:= i_stBms.bComm AND i_stBms.bContactorClosed;
bOpened		:= i_stBms.bComm AND NOT i_stBms.bContactorClosed;
_rtReset(CLK := i_bReset);
_rtWantClose(CLK := i_bWantClose);
CASE i_eProtAction OF
	E_BatAction.Stop:	eProtCmd := E_BatCmd.Open;
	E_BatAction.EStop:	eProtCmd := E_BatCmd.EStop;
ELSE
	eProtCmd := E_BatCmd.None;
END_CASE
IF eProtCmd = E_BatCmd.None THEN
	_bProtNoComm := FALSE;
ELSIF NOT i_stBms.bComm THEN
	_bProtNoComm := TRUE;
END_IF
// 실패 표시 지우기: 투입 요청, 새 기동, 보호 조치가 바뀌면 (다시 보낼 수 있음)
IF i_bCloseReq OR _rtWantClose.Q OR i_eProtAction <> _eLastProt THEN
	q_eFailCmd := E_BatCmd.None;
END_IF
_eLastProt := i_eProtAction;
IF NOT i_bCmdEnable THEN
	_ePending := E_BatCmd.None;		// 설정 오류: 명령을 만들지 않음
	_tonConfirm(IN := FALSE);
	_bResetReq := FALSE;
ELSE
nSeqBefore := _nCmdSeq;
(* 1) 보낸 명령 확인: 바뀌면 끝. 안 바뀌면 보호 명령만 재시도, 나머지는 실패 알람 *)
IF _ePending <> E_BatCmd.None THEN
	IF (_ePending = E_BatCmd.Close AND q_bClosed) OR (_ePending <> E_BatCmd.Close AND bOpened) THEN
		_ePending	:= E_BatCmd.None;
		_nTries		:= 0;
	ELSE
		IF _ePending = E_BatCmd.Close THEN
			_tonConfirm(IN := TRUE, PT := i_stSet.tConfirm);
		ELSE
			_tonConfirm(IN := TRUE, PT := i_stSet.tOpenRetry);
		END_IF
		IF _ePending = eProtCmd AND NOT _bProtNoComm THEN
			_bRetry := TRUE;		// 보호가 같은 명령을 원하면 재시도로 바꿈
		END_IF
		IF _tonConfirm.Q THEN
			IF _bRetry AND _nTries < i_stSet.nOpenRetry THEN
				IF i_stBms.bComm THEN		// 통신이 끊기면 기다렸다가 이어서 보냄
					M_SendCmdAndStartConfirm(_ePending, TRUE);
				END_IF
			ELSE
				q_eFailCmd	:= _ePending;		// 실패 알람만 (잠그지 않음). 같은 명령은 실패를 지울 때까지 다시 보내지 않음
				_ePending	:= E_BatCmd.None;
			END_IF
		END_IF
	END_IF
END_IF
(* 2) 보내기 *)
IF eProtCmd <> E_BatCmd.None THEN
	// 보호 개방·비상정지: 버스 유닛이 멈춘 뒤 (비상정지도 같음). 보호 중에는 투입하지 않음
	IF q_bClosed AND i_bUnitsStopped AND _ePending <> eProtCmd AND q_eFailCmd <> eProtCmd THEN
		M_SendCmdAndStartConfirm(eProtCmd, NOT _bProtNoComm);
	END_IF
ELSIF i_bOpenReq THEN
	IF q_bClosed AND _ePending <> E_BatCmd.Open AND q_eFailCmd <> E_BatCmd.Open THEN
		M_SendCmdAndStartConfirm(E_BatCmd.Open, FALSE);
	END_IF
ELSIF (i_bWantClose OR i_bCloseReq) AND NOT q_bClosed AND i_bUsable
		AND _ePending = E_BatCmd.None AND q_eFailCmd <> E_BatCmd.Close THEN
	M_SendCmdAndStartConfirm(E_BatCmd.Close, FALSE);
END_IF
(* 3) 고장 리셋: BMS가 고장이면 고장 리셋 명령 1회 (확인·재시도 없음)
   보호가 걸려 있어도 보냄. 단, 이번 스캔에 다른 명령을 보냈거나 개방이 진행 중이면 그게 끝난 뒤 보냄 *)
IF _rtReset.Q THEN
	_bResetReq := TRUE;
END_IF
IF _bResetReq THEN
	IF NOT i_stBms.bComm OR NOT i_stBms.bFault THEN
		_bResetReq := FALSE;		// 리셋할 고장 없음 (또는 통신 없음)
	ELSIF _nCmdSeq = nSeqBefore AND (_ePending = E_BatCmd.None OR _ePending = E_BatCmd.Close) THEN
		_nCmdSeq		:= _nCmdSeq + 1;
		q_stCmd.eCmd	:= E_BatCmd.Reset;
		q_stCmd.nSeq	:= _nCmdSeq;
		_bResetReq		:= FALSE;
	END_IF
END_IF
END_IF		// i_bCmdEnable

METHOD PRIVATE M_SendCmdAndStartConfirm	// 명령 1회 보내고 확인 시작
VAR_INPUT
	i_eCmd		: E_BatCmd;
	i_bRetry	: BOOL;		// 확인되지 않으면 재시도 (보호 명령)
END_VAR
IF i_eCmd = _ePending THEN
	_nTries := _nTries + 1;
ELSE
	_nTries := 0;
END_IF
_nCmdSeq		:= _nCmdSeq + 1;
q_stCmd.eCmd	:= i_eCmd;
q_stCmd.nSeq	:= _nCmdSeq;
_ePending		:= i_eCmd;
_bRetry			:= i_bRetry;
_tonConfirm(IN := FALSE);
END_METHOD

END_FUNCTION_BLOCK

// ---- 10_Core/60_Dispatch/FB_BatRequest.TcPOU
FUNCTION_BLOCK FB_BatRequest		// 배터리 그룹(DC 버스)마다 투입·개방 요청 정리: 지령원 BatClose·BatOpen, 정지 시 개방, 운전원이 연 배터리 유지, 거부 이유
// FB_Sequencer 본체가 유닛 시퀀서 다음, BMS 시퀀서 앞에서 부름 (판단만. 명령은 BMS 시퀀서가 만듦)
// 지령원 BatOpen은 버스 유닛이 모두 정지(또는 통신 끊김)했을 때만 (아니면 UnitRunning). 그렇게 연 배터리는 BatClose 또는 그 버스 유닛의 새 기동 요청까지 자동 투입 안 함
VAR_INPUT
	i_bOpenOnStop	: BOOL;			// 정지하면 배터리 개방 (g_stSeqSet.stBat.bOpenOnStop)
END_VAR
VAR_IN_OUT CONSTANT
	iq_astSrcOut	: ARRAY[1..GVL_PARAM.SOURCE_COUNT] OF ST_SourceOutput;
	iq_astReg		: ARRAY[1..GVL_PARAM.SOURCE_COUNT] OF ST_SourceReg;		// 배터리 요청을 받을 운전 모드 (stStateMode.stBat)
	iq_aeOpMode		: ARRAY[1..GVL_PARAM.UNIT_COUNT] OF E_OpMode;			// 실제 운전 모드
	iq_astUnitCfg	: ARRAY[1..GVL_PARAM.UNIT_COUNT] OF ST_UnitCfg;
	iq_astUnit		: ARRAY[1..GVL_PARAM.UNIT_COUNT] OF ST_UnitState;		// 버스 유닛 정지 확인
	iq_abNewReq		: ARRAY[1..GVL_PARAM.UNIT_COUNT] OF BOOL;		// 이번 스캔에 접수된 지령원 상태 요청 있음
	iq_aeReq		: ARRAY[1..GVL_PARAM.UNIT_COUNT] OF E_PcsCmd;	// 그 요청
	iq_abWantBat	: ARRAY[1..GVL_PARAM.BAT_COUNT] OF BOOL;		// 이번 스캔 배터리 투입이 필요함 (순서 기동 유닛, 유닛 시퀀서 결과)
END_VAR
VAR_OUTPUT
	q_abCloseReq	: ARRAY[1..GVL_PARAM.BAT_COUNT] OF BOOL;		// 지령원 BatClose (이번 스캔)
	q_abOpenReq		: ARRAY[1..GVL_PARAM.BAT_COUNT] OF BOOL;		// 개방 요청 (지령원 BatOpen 또는 정지 시 개방)
	q_abBusStopped	: ARRAY[1..GVL_PARAM.BAT_COUNT] OF BOOL;		// 버스 유닛이 모두 정지 확인 (통신 있고 Stop·Fault). 정지 시 개방 기준
	q_abBusStopOk	: ARRAY[1..GVL_PARAM.BAT_COUNT] OF BOOL;		// 버스 유닛이 모두 정지 또는 통신 끊김. 보호 개방·비상정지와 지령원 BatOpen 기준
	q_abHoldOpen	: ARRAY[1..GVL_PARAM.BAT_COUNT] OF BOOL;		// 지령원 BatOpen으로 연 배터리: 다음 투입 요청까지 자동 투입 안 함
	q_aeRefuse		: ARRAY[1..GVL_PARAM.BAT_COUNT] OF E_SeqRefuse;	// 마지막 요청 거부 이유 (새 요청을 받아들이면 None)
	q_abRefusedNow	: ARRAY[1..GVL_PARAM.BAT_COUNT] OF BOOL;		// 이번 스캔에 요청을 거부함 (1스캔, 로그용)
	q_abReqTaken	: ARRAY[1..GVL_PARAM.SOURCE_COUNT] OF BOOL;		// 지령원의 이번 요청을 받은 배터리 그룹이 있음 (로그용)
END_VAR
VAR_TEMP
	u				: UINT;
	b				: UINT;
	i				: UINT;
	bModeOk			: BOOL;		// 이 지령원의 배터리 요청을 받는가 (버스의 유닛 중 하나라도 등록된 운전 모드)
	abReqNow		: ARRAY[1..GVL_PARAM.BAT_COUNT] OF BOOL;		// 이번 스캔에 지령원 요청을 받음
END_VAR

(* 1) 버스마다: 유닛이 모두 정지했나, 그 버스 유닛의 새 기동 요청이 있나 (운전원이 연 배터리도 다시 투입할 수 있음) *)
FOR b := 1 TO GVL_PARAM.BAT_COUNT DO
	q_abBusStopped[b] := TRUE;
	q_abBusStopOk[b]	:= TRUE;
END_FOR
FOR u := 1 TO GVL_PARAM.UNIT_COUNT DO
	b := iq_astUnitCfg[u].nBatGroup;
	IF b >= 1 AND b <= GVL_PARAM.BAT_COUNT THEN
		IF iq_abNewReq[u] AND (iq_aeReq[u] = E_PcsCmd.Run OR iq_aeReq[u] = E_PcsCmd.Standby) THEN
			q_abHoldOpen[b] := FALSE;
		END_IF
		// 정지 확인은 통신이 있고 Stop·Fault일 때 (통신 끊김·Unknown은 정지로 보지 않음)
		IF NOT (iq_astUnit[u].bComm AND F_IsStopped(iq_astUnit[u].eRunState)) THEN
			q_abBusStopped[b] := FALSE;
		END_IF
		// 보호 개방·지령원 BatOpen: 통신이 끊긴 유닛은 정지를 확인할 수 없어 기다리지 않음
		IF iq_astUnit[u].bComm AND NOT F_IsStopped(iq_astUnit[u].eRunState) THEN
			q_abBusStopOk[b] := FALSE;
		END_IF
	END_IF
END_FOR

(* 2) 지령원 배터리 요청 (stBatReq: 배터리 그룹, 0 = 전부). 개방은 버스 유닛이 모두 정지했을 때만 *)
FOR i := 1 TO GVL_PARAM.SOURCE_COUNT DO
	q_abReqTaken[i] := FALSE;
END_FOR
FOR b := 1 TO GVL_PARAM.BAT_COUNT DO
	q_abCloseReq[b]	:= FALSE;
	abReqNow[b]		:= FALSE;
	q_abOpenReq[b]	:= i_bOpenOnStop AND q_abBusStopped[b] AND NOT iq_abWantBat[b];
	FOR i := 1 TO GVL_PARAM.SOURCE_COUNT DO
		bModeOk := FALSE;
		FOR u := 1 TO GVL_PARAM.UNIT_COUNT DO
			IF iq_astUnitCfg[u].nBatGroup = b AND F_BatCmdAllowed(iq_astReg[i].stStateMode.stBat, iq_astSrcOut[i].stBatReq.eCmd, iq_aeOpMode[u]) THEN
				bModeOk := TRUE;
			END_IF
		END_FOR
		IF iq_astSrcOut[i].bValid AND bModeOk AND (iq_astSrcOut[i].stBatReq.nBatGroup = 0 OR iq_astSrcOut[i].stBatReq.nBatGroup = b) THEN
			q_abReqTaken[i]	:= TRUE;
			abReqNow[b]		:= TRUE;
			q_aeRefuse[b]	:= E_SeqRefuse.None;
			IF iq_astSrcOut[i].stBatReq.eCmd = E_BatCmd.Close THEN
				q_abCloseReq[b]	:= TRUE;
				q_abHoldOpen[b]	:= FALSE;
			ELSIF iq_astSrcOut[i].stBatReq.eCmd = E_BatCmd.Open THEN
				IF q_abBusStopOk[b] THEN
					q_abOpenReq[b]	:= TRUE;
					q_abHoldOpen[b]	:= TRUE;		// 운전원이 연 것: 다음 투입 요청까지 자동 투입 안 함
				ELSE
					q_aeRefuse[b] := E_SeqRefuse.UnitRunning;
				END_IF
			END_IF
		END_IF
	END_FOR
	q_abRefusedNow[b] := abReqNow[b] AND q_aeRefuse[b] <> E_SeqRefuse.None;
END_FOR

END_FUNCTION_BLOCK

// ---- 10_Core/40_Arbitration/F_BatCmdAllowed.TcPOU
FUNCTION F_BatCmdAllowed : BOOL		// 지령원의 배터리 요청을 이 운전 모드에서 받나 (명령마다 등록값)
VAR_INPUT
	i_stSet		: ST_BatCmdMode;
	i_eCmd		: E_BatCmd;
	i_eOpMode	: E_OpMode;
END_VAR

CASE i_eCmd OF
	E_BatCmd.Close:		F_BatCmdAllowed := F_SourceAllowed(i_stSet.eClose, i_eOpMode);
	E_BatCmd.Open:		F_BatCmdAllowed := F_SourceAllowed(i_stSet.eOpen, i_eOpMode);
ELSE
	F_BatCmdAllowed := FALSE;		// None, 지령원이 보내지 않는 명령
END_CASE

END_FUNCTION

// ---- 10_Core/40_Arbitration/FB_PermitEval.TcPOU
FUNCTION_BLOCK FB_PermitEval		// 기동 조건 모듈을 그룹마다 스캔당 한 번 평가 (등록된 모듈이 모두 허가해야 기동. 없으면 허가)
// MAIN에서 fbSequencer.M_Prepare 앞에 부름. 시퀀서가 이 결과로 접수 검사·기동 단계를 진행
VAR_IN_OUT CONSTANT
	iq_astView		: ARRAY[1..GVL_PARAM.GROUP_COUNT] OF ST_GroupView;
	iq_astPermitReg	: ARRAY[1..GVL_PARAM.PERMIT_COUNT] OF ST_ModuleReg;
	iq_abWaitPermit	: ARRAY[1..GVL_PARAM.GROUP_COUNT] OF BOOL;		// 그룹이 기동 조건을 기다리는 중 (fbSequencer.q_abWaitPermit, 지난 스캔)
END_VAR
VAR_IN_OUT
	iq_aipPermit	: ARRAY[1..GVL_PARAM.PERMIT_COUNT] OF I_StartPermit;
END_VAR
VAR_OUTPUT
	q_abPermit		: ARRAY[1..GVL_PARAM.GROUP_COUNT] OF BOOL;		// 그룹 기동 조건
	q_anPermitModule: ARRAY[1..GVL_PARAM.GROUP_COUNT] OF UINT;		// 막은 기동 조건 모듈 (처음 것)
	q_anPermitReason: ARRAY[1..GVL_PARAM.GROUP_COUNT] OF UINT;
END_VAR
VAR_TEMP
	g				: UINT;
	i				: UINT;
	bPermitOk		: BOOL;
END_VAR

FOR g := 1 TO GVL_PARAM.GROUP_COUNT DO
	q_abPermit[g]		:= TRUE;
	q_anPermitModule[g]	:= 0;
	q_anPermitReason[g]	:= 0;
	FOR i := 1 TO GVL_PARAM.PERMIT_COUNT DO
		IF iq_aipPermit[i] <> 0 AND_THEN (iq_astPermitReg[i].bEnable
			AND (iq_astPermitReg[i].nGroup = 0 OR iq_astPermitReg[i].nGroup = g)) THEN
			bPermitOk := iq_aipPermit[i].M_Evaluate(i_stView := iq_astView[g], i_bRequest := iq_abWaitPermit[g]);
			IF NOT bPermitOk AND q_abPermit[g] THEN
				q_abPermit[g]		:= FALSE;
				q_anPermitModule[g]	:= iq_aipPermit[i].ModuleId;
				q_anPermitReason[g]	:= iq_aipPermit[i].Reason;
			END_IF
		END_IF
	END_FOR
END_FOR

END_FUNCTION_BLOCK

// ---- 10_Core/60_Dispatch/FB_GroupState.TcPOU
FUNCTION_BLOCK FB_GroupState		// 그룹 상태 요약: 유닛 시퀀스 상태 → 그룹 상태 (그룹 보기에 다음 스캔부터 들어감)
// 우선순위: 운전 > 기동 중 > Standby > 배터리 투입 중 > 정지 중 > 정지. PMS 시작 첫 스캔은 Init
VAR_IN_OUT CONSTANT
	iq_aeUnitSeq	: ARRAY[1..GVL_PARAM.UNIT_COUNT] OF E_UnitSeq;		// fbSequencer.q_aeUnitSeq
	iq_astUnitCfg	: ARRAY[1..GVL_PARAM.UNIT_COUNT] OF ST_UnitCfg;
END_VAR
VAR_OUTPUT
	q_aeGroupState	: ARRAY[1..GVL_PARAM.GROUP_COUNT] OF E_GroupState;
END_VAR
VAR
	_bInit			: BOOL;
END_VAR
VAR_TEMP
	u				: UINT;
	g				: UINT;
	abRunning		: ARRAY[1..GVL_PARAM.GROUP_COUNT] OF BOOL;
	abStarting		: ARRAY[1..GVL_PARAM.GROUP_COUNT] OF BOOL;
	abStandby		: ARRAY[1..GVL_PARAM.GROUP_COUNT] OF BOOL;
	abBatWait		: ARRAY[1..GVL_PARAM.GROUP_COUNT] OF BOOL;
	abStopping		: ARRAY[1..GVL_PARAM.GROUP_COUNT] OF BOOL;
END_VAR

FOR u := 1 TO GVL_PARAM.UNIT_COUNT DO
	g := iq_astUnitCfg[u].nGroup;
	IF g >= 1 AND g <= GVL_PARAM.GROUP_COUNT THEN
		CASE iq_aeUnitSeq[u] OF
			E_UnitSeq.Running:						abRunning[g] := TRUE;
			E_UnitSeq.ToRun, E_UnitSeq.WaitPermit:	abStarting[g] := TRUE;
			E_UnitSeq.Standby:	abStandby[g] := TRUE;
			E_UnitSeq.WaitBat:						abBatWait[g] := TRUE;
			E_UnitSeq.StopRamp, E_UnitSeq.ToStop:	abStopping[g] := TRUE;
		END_CASE
	END_IF
END_FOR

FOR g := 1 TO GVL_PARAM.GROUP_COUNT DO
	IF NOT _bInit THEN
		q_aeGroupState[g] := E_GroupState.Init;
	ELSIF abRunning[g] THEN
		q_aeGroupState[g] := E_GroupState.Running;
	ELSIF abStarting[g] THEN
		q_aeGroupState[g] := E_GroupState.StartWait;
	ELSIF abStandby[g] THEN
		q_aeGroupState[g] := E_GroupState.PcsStandby;
	ELSIF abBatWait[g] THEN
		q_aeGroupState[g] := E_GroupState.BatConnecting;
	ELSIF abStopping[g] THEN
		q_aeGroupState[g] := E_GroupState.Stopping;
	ELSE
		q_aeGroupState[g] := E_GroupState.Stopped;
	END_IF
END_FOR
_bInit := TRUE;

END_FUNCTION_BLOCK

// ---- 10_Core/60_Dispatch/FB_Dispatcher.TcPOU
FUNCTION_BLOCK FB_Dispatcher		// 장비에 쓰는 유일한 곳. 상태 명령: 새 명령일 때 1회. P·Q: Auto = 쓰기 주기마다, Manual = 명령이 들어온 스캔에 바로 1회
VAR_INPUT
	i_tWritePeriod	: TIME;
	i_bWriteEnable	: BOOL := TRUE;	// FALSE = 설정 오류: 장비에 아무것도 쓰지 않음
END_VAR
VAR_IN_OUT
	iq_aipPcs		: ARRAY[1..GVL_PARAM.PCS_COUNT] OF I_Pcs;
	iq_aipBms		: ARRAY[1..GVL_PARAM.BMS_COUNT] OF I_Bms;
END_VAR
VAR_IN_OUT CONSTANT
	iq_astUnitCfg	: ARRAY[1..GVL_PARAM.UNIT_COUNT] OF ST_UnitCfg;
	iq_astUnitCmd	: ARRAY[1..GVL_PARAM.UNIT_COUNT] OF ST_PcsCmd;
	iq_abOutputReady	: ARRAY[1..GVL_PARAM.UNIT_COUNT] OF BOOL;	// 유닛 출력 가능 (FB_OutputReady). Manual 쓰기 시점(들어감·나옴)에만 씀
	iq_astUnitSet	: ARRAY[1..GVL_PARAM.UNIT_COUNT] OF ST_PQ;
	iq_astBmsCmd	: ARRAY[1..GVL_PARAM.BMS_COUNT] OF ST_BatCmd;
	iq_aeOpMode		: ARRAY[1..GVL_PARAM.UNIT_COUNT] OF E_OpMode;
	iq_abManualNew	: ARRAY[1..GVL_PARAM.UNIT_COUNT] OF BOOL;		// 새 수동 지령 (fbManualGate)
	iq_abManualFollow: ARRAY[1..GVL_PARAM.UNIT_COUNT] OF BOOL;		// 램프 중 또는 제한에 걸림 (fbManualShape, FB_ShapePath)
	iq_abUnitLimited: ARRAY[1..GVL_PARAM.UNIT_COUNT] OF BOOL;		// 유닛 지령이 줄었거나 0으로 묶임 (FB_Distributor.q_abUnitLimited)
END_VAR
VAR_OUTPUT
	q_astWritten	: ARRAY[1..GVL_PARAM.UNIT_COUNT] OF ST_PQ;	// 마지막으로 쓴 지령값 (진단용)
	q_abBadSet		: ARRAY[1..GVL_PARAM.UNIT_COUNT] OF BOOL;		// 이번 스캔 지령값이 NaN·무한대여서 0으로 바꿈 (앞 단계 계산 이상)
	q_nBadSetCount	: UDINT;										// 0으로 바꾼 횟수 (PLC 시작 후, 스캔 단위)
END_VAR
VAR
	_anSentUnit		: ARRAY[1..GVL_PARAM.UNIT_COUNT] OF UDINT;	// 보낸 명령 번호
	_anSentBms		: ARRAY[1..GVL_PARAM.BMS_COUNT] OF UDINT;
	_tonWrite		: TON;
	_bStarted		: BOOL;
	_aeLastMode		: ARRAY[1..GVL_PARAM.UNIT_COUNT] OF E_OpMode;
	_abLastReady	: ARRAY[1..GVL_PARAM.UNIT_COUNT] OF BOOL;
	_abFollowing	: ARRAY[1..GVL_PARAM.UNIT_COUNT] OF BOOL;		// 램프·제한을 따라 쓰는 중 (풀린 값까지 쓰면 끝)
END_VAR
VAR_TEMP
	u				: UINT;
	m				: UINT;
	nPcs			: UINT;
	bWrite			: BOOL;
	bWriteNow				: BOOL;
	bFollow			: BOOL;
	bSame			: BOOL;
	stSet			: ST_PQ;
	stZero			: ST_PQ;
END_VAR

_tonWrite(IN := TRUE, PT := i_tWritePeriod);
bWrite := _tonWrite.Q;
IF bWrite THEN
	_tonWrite(IN := FALSE);
END_IF

// PMS 시작 첫 스캔: 수동 유닛은 아무것도 쓰지 않음 (재기동이 운전 중 장비 출력을 바꾸지 않게)
IF NOT _bStarted THEN
	_aeLastMode		:= iq_aeOpMode;
	_abLastReady	:= iq_abOutputReady;
	_bStarted		:= TRUE;
END_IF

FOR u := 1 TO GVL_PARAM.UNIT_COUNT DO
	nPcs := iq_astUnitCfg[u].nPcs;
	IF nPcs >= 1 AND nPcs <= GVL_PARAM.PCS_COUNT AND_THEN iq_aipPcs[nPcs] <> 0 THEN
		// 상태 명령: 새 명령일 때 1회 (Auto·Manual 같음)
		IF iq_astUnitCmd[u].nSeq <> _anSentUnit[u] THEN
			IF iq_astUnitCmd[u].eCmd <> E_PcsCmd.None AND i_bWriteEnable THEN		// 막힌 동안의 명령은 보내지 않고 버림
				iq_aipPcs[nPcs].M_SetStateCmd(i_nSub := iq_astUnitCfg[u].nSub, i_stCmd := iq_astUnitCmd[u]);
			END_IF
			_anSentUnit[u] := iq_astUnitCmd[u].nSeq;
		END_IF

		// 지령값 (출력 못 내는 유닛은 분배에서 이미 0)
		stSet := iq_astUnitSet[u];
		// 마지막 안전장치: NaN·무한대는 장비에 보내지 않고 0 (코어는 실수 계산이라 앞 단계 이상값이 여기까지 올 수 있음)
		q_abBadSet[u] := NOT F_CmdOk(stSet.fP, 0.0) OR NOT F_CmdOk(stSet.fQ, 0.0);
		IF q_abBadSet[u] THEN
			stSet			:= stZero;
			q_nBadSetCount	:= q_nBadSetCount + 1;
		END_IF
		bSame := stSet.fP = q_astWritten[u].fP AND stSet.fQ = q_astWritten[u].fQ;

		IF iq_aeOpMode[u] = E_OpMode.Auto THEN
			(* Auto: 쓰기 주기마다 *)
			bWriteNow := bWrite;
			_abFollowing[u] := FALSE;
		ELSE
			(* Manual: 명령이 들어온 스캔에 바로 1회.
			   그 뒤로는 램프 중이거나 설비 제한(정격·배터리·Derate·제한 모듈)에 걸려 값이 바뀔 때만 쓰기 주기마다 *)
			bFollow := iq_abManualFollow[u]
				OR iq_abUnitLimited[u];
			bWriteNow := iq_abManualNew[u]
				OR iq_aeOpMode[u] <> _aeLastMode[u]				// Auto → Manual 바뀐 스캔
				OR iq_abOutputReady[u] <> _abLastReady[u]	// 출력 가능 들어감·나옴
				OR (bWrite AND (bFollow OR _abFollowing[u]) AND NOT bSame);
			IF bFollow THEN
				_abFollowing[u] := TRUE;
			ELSIF bWriteNow OR bSame THEN
				_abFollowing[u] := FALSE;						// 제한이 풀린 값까지 썼음
			END_IF
		END_IF

		IF bWriteNow AND i_bWriteEnable THEN
			q_astWritten[u] := stSet;
			iq_aipPcs[nPcs].M_SetPower(i_nSub := iq_astUnitCfg[u].nSub, i_fP := stSet.fP, i_fQ := stSet.fQ);
		END_IF
	END_IF
	_aeLastMode[u]		:= iq_aeOpMode[u];
	_abLastReady[u]	:= iq_abOutputReady[u];
END_FOR

FOR m := 1 TO GVL_PARAM.BMS_COUNT DO
	IF iq_aipBms[m] <> 0 AND iq_astBmsCmd[m].nSeq <> _anSentBms[m] THEN
		IF iq_astBmsCmd[m].eCmd <> E_BatCmd.None AND i_bWriteEnable THEN
			iq_aipBms[m].M_SetStateCmd(i_stCmd := iq_astBmsCmd[m]);
		END_IF
		_anSentBms[m] := iq_astBmsCmd[m].nSeq;
	END_IF
END_FOR

END_FUNCTION_BLOCK

// ---- 10_Core/60_Dispatch/FB_AuxOutput.TcPOU
FUNCTION_BLOCK FB_AuxOutput		// 보조 장비 출력(DO)에 쓰는 유일한 곳: 출력 규칙 → 지연·유지 → 같은 점은 OR해서 한 번만 씀
VAR_INPUT
	i_bReset		: BOOL;			// 유지(bLatch) 출력 풀기 (MAIN bClearHoldDo)
	i_bWriteEnable	: BOOL := TRUE;	// FALSE = 설정 오류: DO에 쓰지 않음
END_VAR
VAR_IN_OUT CONSTANT
	iq_astCfg		: ARRAY[1..GVL_PARAM.OUTPUT_COUNT] OF ST_OutputCfg;
END_VAR
VAR_IN_OUT
	iq_aipRule		: ARRAY[1..GVL_PARAM.OUTPUT_COUNT] OF I_OutputRule;
	iq_aipAux		: ARRAY[1..GVL_PARAM.AUX_COUNT] OF I_AuxDevice;
END_VAR
VAR_OUTPUT
	q_abCond		: ARRAY[1..GVL_PARAM.OUTPUT_COUNT] OF BOOL;		// 규칙 판단 (지연 전)
	q_abOn			: ARRAY[1..GVL_PARAM.OUTPUT_COUNT] OF BOOL;		// 이 규칙의 출력 (지연·유지 후)
END_VAR
VAR
	_atonOn			: ARRAY[1..GVL_PARAM.OUTPUT_COUNT] OF TON;
	_atofOff		: ARRAY[1..GVL_PARAM.OUTPUT_COUNT] OF TOF;
	_abLatched		: ARRAY[1..GVL_PARAM.OUTPUT_COUNT] OF BOOL;
	_abPointOut		: ARRAY[1..GVL_PARAM.OUTPUT_COUNT] OF BOOL;		// 이 칸의 점에 쓸 값 (같은 점 규칙 OR, 진단. 쓰기 허가가 없으면 계산만 하고 안 씀)
END_VAR
VAR_TEMP
	i				: UINT;
	k				: UINT;
	nAux			: UINT;
	bFirst			: BOOL;
END_VAR

(* 1) 규칙마다: 판단 → 켜짐 지연 → 꺼짐 지연 → 유지 *)
FOR i := 1 TO GVL_PARAM.OUTPUT_COUNT DO
	q_abCond[i] := FALSE;
	IF iq_aipRule[i] <> 0 AND_THEN iq_astCfg[i].bEnable THEN
		q_abCond[i] := iq_aipRule[i].M_Check(iq_astCfg[i].fThreshold);
	END_IF
	_atonOn[i](IN := q_abCond[i], PT := iq_astCfg[i].tOnDelay);
	_atofOff[i](IN := _atonOn[i].Q, PT := iq_astCfg[i].tOffDelay);

	IF _atonOn[i].Q AND iq_astCfg[i].bLatch THEN
		_abLatched[i] := TRUE;
	END_IF
	IF (i_bReset AND NOT _atonOn[i].Q) OR NOT iq_astCfg[i].bEnable OR NOT iq_astCfg[i].bLatch THEN
		_abLatched[i] := FALSE;
	END_IF
	q_abOn[i] := _atofOff[i].Q OR _abLatched[i];
END_FOR

(* 2) 같은 장비·점에 걸린 규칙은 OR. 점마다 첫 칸에서 한 번만 씀 *)
FOR i := 1 TO GVL_PARAM.OUTPUT_COUNT DO
	_abPointOut[i] := FALSE;
	nAux := iq_astCfg[i].nAux;
	IF nAux >= 1 AND nAux <= GVL_PARAM.AUX_COUNT AND iq_astCfg[i].nPoint >= 1 AND_THEN iq_aipAux[nAux] <> 0 THEN
		bFirst := TRUE;
		FOR k := 1 TO GVL_PARAM.OUTPUT_COUNT DO
			IF iq_astCfg[k].nAux = nAux AND iq_astCfg[k].nPoint = iq_astCfg[i].nPoint THEN
				_abPointOut[i] := _abPointOut[i] OR q_abOn[k];
				IF k < i THEN
					bFirst := FALSE;
				END_IF
			END_IF
		END_FOR
		// 쓰기 허가가 없으면(설정 오류·대기 PLC) 켜는 쓰기만 막고 끄는 쓰기는 함: 펄스 출력(차단기 코일 등)이 켜진 채 남지 않게
		IF bFirst AND (i_bWriteEnable OR NOT _abPointOut[i]) THEN
			iq_aipAux[nAux].M_SetBit(i_nPoint := iq_astCfg[i].nPoint, i_bValue := _abPointOut[i]);
		END_IF
	END_IF
END_FOR

END_FUNCTION_BLOCK

// ---- 10_Core/70_Diag/FB_OutputDiag.TcPOU
FUNCTION_BLOCK FB_OutputDiag		// 그룹마다 출력을 처음 막은 단계·주체·이유 (매 스캔). 경로(Auto/Manual)·P/Q별로 4개. 두 경로가 같은 방식
// 이벤트 로그(출력 제한·해소)와 보고는 Auto P(q_astAutoPDiag)만 씀
VAR_IN_OUT CONSTANT
	iq_astAutoShape		: ARRAY[1..GVL_PARAM.GROUP_COUNT] OF ST_ShapeDiag;
	iq_astManualShape	: ARRAY[1..GVL_PARAM.GROUP_COUNT] OF ST_ShapeDiag;
	iq_astDist			: ARRAY[1..GVL_PARAM.GROUP_COUNT] OF ST_DistDiag;
	iq_astUnitDiag		: ARRAY[1..GVL_PARAM.UNIT_COUNT] OF ST_UnitDiag;
	iq_aeOpMode			: ARRAY[1..GVL_PARAM.UNIT_COUNT] OF E_OpMode;
	iq_aeGroupState		: ARRAY[1..GVL_PARAM.GROUP_COUNT] OF E_GroupState;
	iq_astWritten		: ARRAY[1..GVL_PARAM.UNIT_COUNT] OF ST_PQ;
	iq_astUnitSet		: ARRAY[1..GVL_PARAM.UNIT_COUNT] OF ST_PQ;		// 분배 결과 (추적표용)
	iq_astUnitCfg		: ARRAY[1..GVL_PARAM.UNIT_COUNT] OF ST_UnitCfg;
END_VAR
VAR_OUTPUT
	q_astAutoPDiag		: ARRAY[1..GVL_PARAM.GROUP_COUNT] OF ST_OutputDiag;		// Auto 유닛 P (kW). 이벤트 로그·보고는 이것만 씀
	q_astManualPDiag	: ARRAY[1..GVL_PARAM.GROUP_COUNT] OF ST_OutputDiag;		// Manual 유닛 P (kW)
	q_astAutoQDiag		: ARRAY[1..GVL_PARAM.GROUP_COUNT] OF ST_OutputDiag;		// Auto 유닛 Q (kvar)
	q_astManualQDiag	: ARRAY[1..GVL_PARAM.GROUP_COUNT] OF ST_OutputDiag;		// Manual 유닛 Q (kvar)
	q_astAutoPTrace		: ARRAY[1..GVL_PARAM.GROUP_COUNT] OF ST_PTrace;		// Auto P 추적표: 요청 → … → 쓴 값 (접속점 기준이라 그룹 전체 유닛 합)
	q_astManualPTrace	: ARRAY[1..GVL_PARAM.GROUP_COUNT] OF ST_PTrace;		// Manual P 추적표: 요청 → … → 쓴 값 (Manual 유닛 합)
END_VAR
VAR_TEMP
	g				: UINT;
	u				: UINT;
	nAutoUnits		: UINT;
	nManualUnits	: UINT;
	eAutoPBy		: E_UnitLimitBy;	// 그룹 안 그 경로 유닛 중 처음 찾은 제한 이유
	eManualPBy			: E_UnitLimitBy;
	eAutoQBy		: E_UnitLimitBy;
	eManualQBy			: E_UnitLimitBy;
	fAllSet			: REAL;			// 분배 후 그룹 전체 유닛 P 합
	fAllWritten		: REAL;			// 장비에 쓴 그룹 전체 유닛 P 합
	fManualSet			: REAL;			// 분배 후 Manual 유닛 P 합
	fManualWritten		: REAL;
END_VAR

FOR g := 1 TO GVL_PARAM.GROUP_COUNT DO
	q_astAutoPDiag[g]	:= M_Clear(iq_aeGroupState[g]);
	q_astManualPDiag[g]	:= M_Clear(iq_aeGroupState[g]);
	q_astAutoQDiag[g]	:= M_Clear(iq_aeGroupState[g]);
	q_astManualQDiag[g]	:= M_Clear(iq_aeGroupState[g]);
	nAutoUnits		:= 0;
	nManualUnits	:= 0;
	eAutoPBy		:= E_UnitLimitBy.None;
	eManualPBy			:= E_UnitLimitBy.None;
	eAutoQBy		:= E_UnitLimitBy.None;
	eManualQBy			:= E_UnitLimitBy.None;
	fAllSet			:= 0;
	fAllWritten		:= 0;
	fManualSet			:= 0;
	fManualWritten		:= 0;

	// 경로별 유닛 수와 쓴 값 합 (각 진단은 그 경로 유닛만)
	FOR u := 1 TO GVL_PARAM.UNIT_COUNT DO
		IF iq_astUnitCfg[u].nGroup = g THEN
			fAllSet		:= fAllSet + iq_astUnitSet[u].fP;
			fAllWritten	:= fAllWritten + iq_astWritten[u].fP;
			IF iq_aeOpMode[u] = E_OpMode.Manual THEN
				nManualUnits				:= nManualUnits + 1;
				fManualSet						:= fManualSet + iq_astUnitSet[u].fP;
				fManualWritten					:= fManualWritten + iq_astWritten[u].fP;
				q_astManualPDiag[g].fOut	:= q_astManualPDiag[g].fOut + iq_astWritten[u].fP;
				q_astManualQDiag[g].fOut	:= q_astManualQDiag[g].fOut + iq_astWritten[u].fQ;
				M_FirstBy(iq_eBy := eManualPBy, i_eUnitBy := iq_astUnitDiag[u].ePBy);
				M_FirstBy(iq_eBy := eManualQBy, i_eUnitBy := iq_astUnitDiag[u].eQBy);
			ELSE
				nAutoUnits					:= nAutoUnits + 1;
				q_astAutoPDiag[g].fOut		:= q_astAutoPDiag[g].fOut + iq_astWritten[u].fP;
				q_astAutoQDiag[g].fOut		:= q_astAutoQDiag[g].fOut + iq_astWritten[u].fQ;
				M_FirstBy(iq_eBy := eAutoPBy, i_eUnitBy := iq_astUnitDiag[u].ePBy);
				M_FirstBy(iq_eBy := eAutoQBy, i_eUnitBy := iq_astUnitDiag[u].eQBy);
			END_IF
		END_IF
	END_FOR

	// 추적표: 성형이 만든 줄 뒤에 유닛 한도·분배 후 합, 쓴 값 합을 덧붙임
	q_astAutoPTrace[g]		:= M_AddUnitSteps(i_stTrace := iq_astAutoShape[g].stTrace, i_fUnitSum := fAllSet, i_fWritten := fAllWritten);
	q_astManualPTrace[g]	:= M_AddUnitSteps(i_stTrace := iq_astManualShape[g].stTrace, i_fUnitSum := fManualSet, i_fWritten := fManualWritten);

	// P: 요청 → 이 경로 유닛 → 그룹 운전 → 최종 값을 정한 곳 (추적표에서 값을 바꾼 마지막 단계)
	M_StageP(iq_stDiag := q_astAutoPDiag[g], i_stShape := iq_astAutoShape[g], i_stTrace := q_astAutoPTrace[g], i_eUnitBy := eAutoPBy, i_nUnits := nAutoUnits);
	M_StageP(iq_stDiag := q_astManualPDiag[g], i_stShape := iq_astManualShape[g], i_stTrace := q_astManualPTrace[g], i_eUnitBy := eManualPBy, i_nUnits := nManualUnits);
	// Manual P: 추적표에서 값이 안 바뀌었어도 Manual 유닛이 유닛 한도에 걸렸으면 표시 (Manual 진단은 처음 막은 곳)
	IF q_astManualPDiag[g].eStage = E_DiagStage.None AND eManualPBy <> E_UnitLimitBy.None THEN
		q_astManualPDiag[g].eStage	:= E_DiagStage.UnitLimit;
		q_astManualPDiag[g].eUnitBy	:= eManualPBy;
	END_IF

	// Q: 요청 → 이 경로 유닛 → 그룹 운전 → 설비 제한 → 유닛 한도·분배 (UnitLimit 이유는 eUnitBy, 분배 축소만이면 None)
	M_StageQ(iq_stDiag := q_astAutoQDiag[g], i_stShape := iq_astAutoShape[g], i_stDist := iq_astDist[g].stAutoQ, i_eUnitBy := eAutoQBy, i_nUnits := nAutoUnits);
	M_StageQ(iq_stDiag := q_astManualQDiag[g], i_stShape := iq_astManualShape[g], i_stDist := iq_astDist[g].stManualQ, i_eUnitBy := eManualQBy, i_nUnits := nManualUnits);
END_FOR

METHOD PRIVATE M_Clear : ST_OutputDiag		// 빈 진단 + 그룹 상태
VAR_INPUT
	i_eState	: E_GroupState;
END_VAR
VAR
	stNone		: ST_OutputDiag;
END_VAR
M_Clear := stNone;
M_Clear.eGroupState := i_eState;
END_METHOD

METHOD PRIVATE M_FirstBy		// 처음 찾은 유닛 제한 이유만 남김 (모드 전환은 제외)
VAR_IN_OUT
	iq_eBy		: E_UnitLimitBy;
END_VAR
VAR_INPUT
	i_eUnitBy	: E_UnitLimitBy;
END_VAR
IF iq_eBy = E_UnitLimitBy.None AND i_eUnitBy <> E_UnitLimitBy.ModeSwitch THEN
	iq_eBy := i_eUnitBy;
END_IF
END_METHOD

METHOD PRIVATE M_AddUnitSteps : ST_PTrace		// 추적표 끝에 분배 후 합·쓴 값 합 두 줄
VAR_INPUT
	i_stTrace	: ST_PTrace;
	i_fUnitSum	: REAL;
	i_fWritten	: REAL;
END_VAR
M_AddUnitSteps := i_stTrace;
IF M_AddUnitSteps.nCount >= 1 AND M_AddUnitSteps.nCount <= GVL_PARAM.TRACE_STEP_MAX - 2 THEN
	M_AddUnitSteps.nCount := M_AddUnitSteps.nCount + 1;
	M_AddUnitSteps.astStep[M_AddUnitSteps.nCount].eStep		:= E_TraceStep.UnitDist;
	M_AddUnitSteps.astStep[M_AddUnitSteps.nCount].fValue	:= i_fUnitSum;
	M_AddUnitSteps.astStep[M_AddUnitSteps.nCount].bCut		:= ABS(i_fUnitSum - M_AddUnitSteps.astStep[M_AddUnitSteps.nCount - 1].fValue) > 1.0;
	M_AddUnitSteps.nCount := M_AddUnitSteps.nCount + 1;
	M_AddUnitSteps.astStep[M_AddUnitSteps.nCount].eStep		:= E_TraceStep.Written;
	M_AddUnitSteps.astStep[M_AddUnitSteps.nCount].fValue	:= i_fWritten;
END_IF
END_METHOD

METHOD PRIVATE M_StageP		// P 진단: 요청 → 유닛 → 운전 → 추적표에서 값을 바꾼 마지막 단계
VAR_IN_OUT
	iq_stDiag	: ST_OutputDiag;
END_VAR
VAR_INPUT
	i_stShape	: ST_ShapeDiag;
	i_stTrace	: ST_PTrace;
	i_eUnitBy	: E_UnitLimitBy;	// 그 경로 유닛 중 처음 찾은 유닛 한도 이유
	i_nUnits	: UINT;
END_VAR
VAR
	k			: INT;
END_VAR
iq_stDiag.fReq := i_stShape.fPReq;		// 그룹 지령 또는 유닛 지령 합
IF NOT i_stShape.bPGroupCmd AND NOT i_stShape.bPUnitCmd THEN
	iq_stDiag.eStage := E_DiagStage.NoRequest;
ELSIF i_nUnits = 0 THEN
	iq_stDiag.eStage := E_DiagStage.NoUnit;
ELSIF iq_stDiag.eGroupState <> E_GroupState.Running THEN
	iq_stDiag.eStage := E_DiagStage.NotRunning;
ELSE
	FOR k := TO_INT(i_stTrace.nCount) TO 1 BY -1 DO
		IF iq_stDiag.eStage = E_DiagStage.None AND i_stTrace.astStep[k].bCut THEN
			CASE i_stTrace.astStep[k].eStep OF
				E_TraceStep.Ramp:		iq_stDiag.eStage := E_DiagStage.Ramp;
				E_TraceStep.PccLimit:	iq_stDiag.eStage := E_DiagStage.PccLimit;
				E_TraceStep.DevRating, E_TraceStep.DevBattery, E_TraceStep.DevLimit:
										iq_stDiag.eStage := E_DiagStage.DeviceLimit;
				E_TraceStep.UnitDist:	iq_stDiag.eStage := E_DiagStage.UnitLimit;
			END_CASE
			IF iq_stDiag.eStage = E_DiagStage.UnitLimit THEN
				iq_stDiag.eUnitBy	:= i_eUnitBy;		// 유닛 한도 이유 (분배 축소만이면 None)
			ELSIF iq_stDiag.eStage <> E_DiagStage.None THEN
				iq_stDiag.nModule	:= i_stTrace.astStep[k].nModule;
				iq_stDiag.nReason	:= i_stTrace.astStep[k].nReason;
			END_IF
		END_IF
	END_FOR
END_IF
END_METHOD

METHOD PRIVATE M_StageQ		// Q 진단: 요청 → 유닛 → 운전 → 설비 제한 → 유닛 한도·분배 (Q는 램프 없음)
VAR_IN_OUT
	iq_stDiag	: ST_OutputDiag;
END_VAR
VAR_INPUT
	i_stShape	: ST_ShapeDiag;
	i_stDist	: ST_DistPathDiag;
	i_eUnitBy	: E_UnitLimitBy;
	i_nUnits	: UINT;
END_VAR
iq_stDiag.fReq := i_stShape.stQ.fIn;
IF NOT i_stShape.bQGroupCmd AND NOT i_stShape.bQUnitCmd THEN
	iq_stDiag.eStage := E_DiagStage.NoRequest;
ELSIF i_nUnits = 0 THEN
	iq_stDiag.eStage := E_DiagStage.NoUnit;
ELSIF iq_stDiag.eGroupState <> E_GroupState.Running THEN
	iq_stDiag.eStage := E_DiagStage.NotRunning;
ELSIF i_stShape.stQ.bClamped THEN
	iq_stDiag.eStage	:= E_DiagStage.DeviceLimit;
	iq_stDiag.nModule	:= i_stShape.stQ.nModule;
	iq_stDiag.nReason	:= i_stShape.stQ.nReason;
ELSIF ABS(i_stDist.fShareReq - i_stDist.fShareGot) > 1.0 OR i_stDist.fFixedScale < 0.999 OR i_eUnitBy <> E_UnitLimitBy.None THEN
	iq_stDiag.eStage	:= E_DiagStage.UnitLimit;
	iq_stDiag.eUnitBy	:= i_eUnitBy;
END_IF
END_METHOD

END_FUNCTION_BLOCK

// ---- 10_Core/70_Diag/FB_EventLog.TcPOU
FUNCTION_BLOCK FB_EventLog		// 기록하는 유일한 곳: 결과를 보고 바뀔 때만 이벤트 로거에 남김
VAR_INPUT
	i_stSet			: ST_LogSet;
	i_bTestMode		: BOOL;			// 시험 모드에서만 가상신호를 씀 (가상신호 알람도)
	i_bSetChanged	: BOOL;			// 운영 설정이 바뀌어 저장 시작 (FB_PersistSave.q_bSetChanged, 1스캔)
	i_sSetChanged	: WSTRING(63);	// 바뀐 설정 이름
	i_bSetRejected	: BOOL;			// 잘못된 설정 값을 마지막 정상값으로 되돌림 (FB_SettingGuard.q_bRejected, 1스캔)
	i_sSetRejected	: WSTRING(63);	// 되돌린 설정과 이유
	i_bPersistError	: BOOL;			// 설정 저장 실패 (FB_PersistSave.q_bError)
	i_nPersistErrorId	: UDINT;	// 그 오류 번호
	i_nConfigErrors	: UINT;			// 설정 오류 수 (FB_ConfigCheck.q_nErrors)
	i_bPmsStart		: BOOL;			// PMS 시작 (FB_AliveRecorder.q_bStartEvent, 1스캔)
	i_sStartLastAlive	: WSTRING(63);	// 직전 동작 시각 (글자)
	i_sStartOffTime	: WSTRING(63);	// 꺼져 있던 시간 (글자)
	(* 이중화 (GVL_IF) *)
	i_bRedUse		: BOOL;			// 이중화를 씀 (GVL_SITE.RED_SET.bUse)
	i_eRedRole		: E_RedRole;
	i_eRedState		: E_RedState;
	i_ePeer			: E_RedPeer;
	i_nSwitchCount	: UDINT;		// Active가 바뀐 횟수 (GVL_IF.g_nRedSwitchCount)
	i_eSwitch		: E_RedSwitch;	// 마지막으로 바뀐 이유
	i_nResumeCount	: UDINT;		// PLC가 멈췄다 이어진 횟수
	i_nSyncApplied	: UDINT;		// 상대 값으로 설정을 덮어쓴 횟수
	i_bSyncFresh	: BOOL;			// 상대의 동기화 값이 낡지 않음
	i_bPeerEapOk	: BOOL;
	i_bRoleConflict	: BOOL;			// 두 PLC 역할이 같음
	(* MQTT 브로커 끊김 (FB_BrokerWatch) [9번 수정 2026-11-09: 추가] *)
	i_bBrokerLost	: BOOL;			// 고른 브로커가 판정 시간 넘게 끊김 (알람)
	i_sBrokerName	: WSTRING(15);	// 브로커 이름 (Cloud·Local·Azure)
	i_sBrokerDelay	: WSTRING(31);	// 판정 시간 (글자)
END_VAR
VAR_IN_OUT CONSTANT
	iq_asConfigErrors	: ARRAY[1..10] OF WSTRING(63);	// 설정 오류 문구 (FB_ConfigCheck.q_asErrors)
	(* 보호 *)
	iq_aabRule		: ARRAY[1..GVL_PARAM.RULE_COUNT, 1..GVL_PARAM.PROT_TARGET_MAX] OF BOOL;	// 보호 발생 [규칙 칸, 대상] (FB_Protection.q_aabRule)
	iq_astRuleCfg	: ARRAY[1..GVL_PARAM.RULE_COUNT] OF ST_RuleCfg;
	(* 시퀀스 *)
	iq_aeUnitSeq	: ARRAY[1..GVL_PARAM.UNIT_COUNT] OF E_UnitSeq;
	iq_aeRefuse		: ARRAY[1..GVL_PARAM.UNIT_COUNT] OF E_SeqRefuse;
	iq_aeBatRefuse	: ARRAY[1..GVL_PARAM.BAT_COUNT] OF E_SeqRefuse;	// 배터리 그룹별 요청 거부 이유
	iq_abBatRefusedNow: ARRAY[1..GVL_PARAM.BAT_COUNT] OF BOOL;		// 이번 스캔에 배터리 요청 거부
	iq_aeFailCmd	: ARRAY[1..GVL_PARAM.UNIT_COUNT] OF E_PcsCmd;
	iq_aeBmsFailCmd	: ARRAY[1..GVL_PARAM.BMS_COUNT] OF E_BatCmd;	// 확인되지 않은 BMS 명령 (FB_Sequencer)
	iq_aeOpMode		: ARRAY[1..GVL_PARAM.UNIT_COUNT] OF E_OpMode;
	iq_abModeForced	: ARRAY[1..GVL_PARAM.UNIT_COUNT] OF BOOL;		// 보호가 요청 모드를 Manual로 바꾼 스캔 (FB_ModeSwitch.q_abModeForced, 1스캔)
	iq_astUnitProt	: ARRAY[1..GVL_PARAM.UNIT_COUNT] OF ST_UnitProt;	// 보호 결과 (모드 조치를 건 주체 이름)
	(* 명령 필터 *)
	iq_abBadValue	: ARRAY[1..GVL_PARAM.SOURCE_COUNT] OF BOOL;
	iq_afBadValue	: ARRAY[1..GVL_PARAM.SOURCE_COUNT] OF REAL;
	iq_aeManualRefuse	: ARRAY[1..GVL_PARAM.UNIT_COUNT] OF E_CmdRefuse;
	iq_anManualRefuseModule: ARRAY[1..GVL_PARAM.UNIT_COUNT] OF UINT;
	(* 지령원 *)
	iq_astSrcOut	: ARRAY[1..GVL_PARAM.SOURCE_COUNT] OF ST_SourceOutput;
	iq_abPcsReqTaken: ARRAY[1..GVL_PARAM.SOURCE_COUNT] OF BOOL;
	iq_abBatReqTaken: ARRAY[1..GVL_PARAM.SOURCE_COUNT] OF BOOL;		// 시퀀서가 받은 배터리 요청
	iq_astReg		: ARRAY[1..GVL_PARAM.SOURCE_COUNT] OF ST_SourceReg;
	(* 출력 *)
	iq_astAutoPDiag	: ARRAY[1..GVL_PARAM.GROUP_COUNT] OF ST_OutputDiag;
	iq_astUnitDiag	: ARRAY[1..GVL_PARAM.UNIT_COUNT] OF ST_UnitDiag;
	iq_astVirtual	: ARRAY[1..GVL_PARAM.GROUP_COUNT] OF ST_VirtualSet;
	iq_abBadSet		: ARRAY[1..GVL_PARAM.UNIT_COUNT] OF BOOL;		// 지령값 NaN·무한대 → 0 (FB_Dispatcher.q_abBadSet)
	(* 기동 조건 *)
	iq_abWaitPermit	: ARRAY[1..GVL_PARAM.GROUP_COUNT] OF BOOL;		// 기동 조건 기다리는 중 (FB_Sequencer.q_abWaitPermit)
	iq_abPermit		: ARRAY[1..GVL_PARAM.GROUP_COUNT] OF BOOL;		// 기동 조건 (FB_PermitEval)
	iq_anPermitModule: ARRAY[1..GVL_PARAM.GROUP_COUNT] OF UINT;		// 막은 모듈
	iq_anPermitReason: ARRAY[1..GVL_PARAM.GROUP_COUNT] OF UINT;
	(* 장비 상태 (쓰기 실패) *)
	iq_astUnit		: ARRAY[1..GVL_PARAM.UNIT_COUNT] OF ST_UnitState;	// FB_Snapshot.q_astUnit
	iq_astBms		: ARRAY[1..GVL_PARAM.BMS_COUNT] OF ST_BatState;		// FB_Snapshot.q_astBms
END_VAR
VAR_IN_OUT
	iq_aipRule		: ARRAY[1..GVL_PARAM.RULE_COUNT] OF I_ProtectionRule;
	iq_aipResp		: ARRAY[1..GVL_PARAM.RULE_COUNT] OF I_ProtResponse;	// [결함 8 수정 2026-11-03: 추가] 보호 대응 (GVL_SITE.g_aipResp). 빈 칸은 조치 없음 → 알람 문구·심각도도 조치 없음으로
	iq_aipSource	: ARRAY[1..GVL_PARAM.SOURCE_COUNT] OF I_CommandSource;
	iq_aipModule	: ARRAY[1..GVL_PARAM.MODULE_MAX] OF I_Module;	// 등록된 모듈 전부 (FB_ModuleList): 이름·이유 문구 찾기
	iq_fbCtrlMode	: FB_CtrlModeMgr;	// 제어 모드 관리자 (GVL_SITE.g_fbCtrlMode1): 켜진 모드 바뀜·요청 거부·스스로 끝남 기록. 관리자를 늘리면 입력도 늘림 [7번 수정 2026-11-09: 추가]
END_VAR
VAR
	(* 알람 *)
	_aafbRule		: ARRAY[1..GVL_PARAM.RULE_COUNT, 1..GVL_PARAM.PROT_TARGET_MAX] OF FB_LogAlarm;	// 보호 [규칙 칸, 대상]
	_afbBmsCmdFail	: ARRAY[1..GVL_PARAM.BMS_COUNT] OF FB_LogAlarm;
	_afbCmdFail		: ARRAY[1..GVL_PARAM.UNIT_COUNT] OF FB_LogAlarm;
	_afbSrcLost		: ARRAY[1..GVL_PARAM.SOURCE_COUNT] OF FB_LogAlarm;
	_afbVirtual		: ARRAY[1..GVL_PARAM.GROUP_COUNT] OF FB_LogAlarm;
	_afbUnitWriteFail	: ARRAY[1..GVL_PARAM.UNIT_COUNT] OF FB_LogAlarm;	// 유닛 쓰기 실패
	_afbBmsWriteFail	: ARRAY[1..GVL_PARAM.BMS_COUNT] OF FB_LogAlarm;		// BMS 쓰기 실패
	_fbPersistFail	: FB_LogAlarm;		// 설정 저장 실패
	_fbControlBlocked	: FB_LogAlarm;	// 설정 오류로 장비 제어 중지
	_fbConfigError	: FB_LogMsg;		// 설정 오류 문구
	_asCfgLogged	: ARRAY[1..10] OF WSTRING(63);	// 마지막으로 기록한 설정 오류 문구
	_nCfgLogged		: UINT;
	_bCfgStarted	: BOOL;
	(* 메시지 *)
	_fbStateReq		: FB_LogMsg;
	_fbLimited		: FB_LogMsg;
	_fbFree			: FB_LogMsg;
	_fbUnitLim		: FB_LogMsg;
	_fbRefused		: FB_LogMsg;
	_fbSeqChange	: FB_LogMsg;
	_fbModeChange	: FB_LogMsg;
	_fbCmdRefused	: FB_LogMsg;
	_fbSetChanged	: FB_LogMsg;		// 운영 설정 바뀜
	_fbSetRejected	: FB_LogMsg;		// 잘못된 설정 값 되돌림
	_fbPermitWait	: FB_LogMsg;		// 기동 조건 대기
	_fbBadSet		: FB_LogMsg;		// 지령값 이상
	_fbPmsStart		: FB_LogMsg;		// PMS 시작
	(* 이중화 *)
	_fbRedStart		: FB_LogMsg;		// Active로 시작
	_fbRedFailover	: FB_LogMsg;		// 절체
	_fbRedFailback	: FB_LogMsg;		// 복귀
	_fbRedYield		: FB_LogMsg;		// Active 양보
	_fbRedResume	: FB_LogMsg;		// 멈췄다 이어짐
	_fbRedSyncApplied: FB_LogMsg;		// 동기화로 설정을 맞춤
	_fbRedPeerLost	: FB_LogAlarm;		// 상대 PLC 끊김
	_fbRedLinkFault	: FB_LogAlarm;		// 통신 한쪽 고장
	_fbRedSyncLost	: FB_LogAlarm;		// 동기화 값을 못 받음
	_fbRedFailed	: FB_LogAlarm;		// 이중화 설정 오류
	_tonRedSync		: TON;
	_tonRedQuiet	: TON;
	_bRedQuiet		: BOOL;				// 멈췄다 이어진 직후: 횟수·이유가 어긋나게 읽힐 수 있어 절체 기록을 잠시 건너뜀
	_bRedInit		: BOOL;
	_bRedSwitchPending: BOOL;
	_nRedSwitchLast	: UDINT;
	_nRedResumeLast	: UDINT;
	_nRedAppliedLast: UDINT;
	_fbModeForced	: FB_LogMsg;		// 보호가 운전 모드를 Manual로 바꿈
	(* [7번 수정 2026-11-09: 추가] 제어 모드 *)
	_fbCmChange		: FB_LogMsg;		// 켜진 제어 모드 바뀜
	_fbCmRefused	: FB_LogMsg;		// 제어 모드 요청 거부
	_fbCmExit		: FB_LogMsg;		// 제어 모드 스스로 끝남
	_nCmLogged		: UINT;				// 마지막으로 기록한 켜진 모드 칸 (0 = 없음)
	_fbBrokerLost	: FB_LogAlarm;		// MQTT 브로커 끊김 [9번 수정 2026-11-09: 추가]
	(* 이전 값 *)
	_aeLastPcsReq	: ARRAY[1..GVL_PARAM.SOURCE_COUNT] OF E_PcsCmd;	// 지령원별 마지막으로 기록한 PCS 요청
	_anLastPcsUnit	: ARRAY[1..GVL_PARAM.SOURCE_COUNT] OF UINT;
	_abEverValid	: ARRAY[1..GVL_PARAM.SOURCE_COUNT] OF BOOL;
	_anVirtualKind	: ARRAY[1..GVL_PARAM.GROUP_COUNT] OF UINT;	// 알람에 올린 가상신호 종류
	_astLogged		: ARRAY[1..GVL_PARAM.GROUP_COUNT] OF ST_OutputDiag;	// 마지막으로 기록한 출력 진단
	_astCand		: ARRAY[1..GVL_PARAM.GROUP_COUNT] OF ST_OutputDiag;	// 유지 시간 재는 중인 후보
	_atonHold		: ARRAY[1..GVL_PARAM.GROUP_COUNT] OF TON;
	_aeLastLimBy	: ARRAY[1..GVL_PARAM.UNIT_COUNT] OF E_UnitLimitBy;
	_aeLastRefuse	: ARRAY[1..GVL_PARAM.UNIT_COUNT] OF E_SeqRefuse;
	_aeLastSeq		: ARRAY[1..GVL_PARAM.UNIT_COUNT] OF E_UnitSeq;
	_aeLastMode		: ARRAY[1..GVL_PARAM.UNIT_COUNT] OF E_OpMode;
	_abLastBad		: ARRAY[1..GVL_PARAM.SOURCE_COUNT] OF BOOL;
	_aeLastCmdRefuse: ARRAY[1..GVL_PARAM.UNIT_COUNT] OF E_CmdRefuse;
	_abPermitLogged	: ARRAY[1..GVL_PARAM.GROUP_COUNT] OF BOOL;	// 이번 대기에서 기동 조건 대기를 기록함
	_anPermitModule	: ARRAY[1..GVL_PARAM.GROUP_COUNT] OF UINT;	// 기록한 막은 모듈·이유 (바뀌면 다시 기록)
	_anPermitReason	: ARRAY[1..GVL_PARAM.GROUP_COUNT] OF UINT;
	_abLastBadSet	: ARRAY[1..GVL_PARAM.UNIT_COUNT] OF BOOL;
	_abModeForcedLogged	: ARRAY[1..GVL_PARAM.UNIT_COUNT] OF BOOL;	// 이번 보호(모드 조치)에서 기록함. 보호가 풀리면 다시 기록 가능 (Auto 재요청을 되돌릴 때마다 남기지 않음)
	_bInit			: BOOL;
	(* 모듈 이름 찾기용 사본 (메서드에서 씀) *)
	_aipModule	: ARRAY[1..GVL_PARAM.MODULE_MAX] OF I_Module;
	(* 반복 변수·임시값: 본문과 기록 액션(A_Log...)이 함께 씀. 액션이 본문의 VAR_TEMP를 못 볼 수 있어 VAR에 둠 *)
	_i				: UINT;
	_g				: UINT;
	_u				: UINT;
	_m				: UINT;
	_t				: UINT;			// 보호 대상 번호
	_dwBadBits		: DWORD;		// 이상값 비트 (NaN 구별). [결함 9 수정 2026-11-03: 추가]
	_stProtTxt		: ST_ProtCfg;	// [결함 8 수정 2026-11-03: 추가] 알람 문구에 쓰는 조치 (대응 칸이 비면 조치 없음)
	_b				: UINT;
	_nVirtualKind	: UINT;		// 가상신호 종류: 0 없음, 1 전압, 2 유효전력, 3 둘 다
	_bLost			: BOOL;
	_bCfgChanged	: BOOL;
	_asArg			: ARRAY[1..6] OF WSTRING(63);
END_VAR

_aipModule := iq_aipModule;

// 이번 스캔 인자 비움 (예전 VAR_TEMP와 같은 동작)
FOR _i := 1 TO 6 DO
	_asArg[_i] := "";
END_FOR

IF NOT _bInit THEN
	FOR _u := 1 TO GVL_PARAM.UNIT_COUNT DO
		_aeLastSeq[_u]	:= iq_aeUnitSeq[_u];
		_aeLastMode[_u]	:= iq_aeOpMode[_u];
	END_FOR
END_IF

_fbStateReq(i_stEntry := TC_EVENTS.PmsSeq.StateRequest);
_fbLimited(i_stEntry := TC_EVENTS.PmsOutput.OutputLimited);
_fbFree(i_stEntry := TC_EVENTS.PmsOutput.OutputFree);
_fbUnitLim(i_stEntry := TC_EVENTS.PmsOutput.UnitLimited);
_fbRefused(i_stEntry := TC_EVENTS.PmsSeq.ReqRefused);
_fbSeqChange(i_stEntry := TC_EVENTS.PmsSeq.SeqChange);
_fbModeChange(i_stEntry := TC_EVENTS.PmsSeq.ModeChange);
_fbCmdRefused(i_stEntry := TC_EVENTS.PmsSeq.CmdRefused);
_fbSetChanged(i_stEntry := TC_EVENTS.PmsSystem.SettingChanged);
_fbConfigError(i_stEntry := TC_EVENTS.PmsSystem.ConfigError);
_fbPermitWait(i_stEntry := TC_EVENTS.PmsSeq.PermitWait);
_fbBadSet(i_stEntry := TC_EVENTS.PmsOutput.BadSetpoint);
_fbPmsStart(i_stEntry := TC_EVENTS.PmsSystem.PmsStart);
_fbRedStart(i_stEntry := TC_EVENTS.PmsSystem.RedStart);
_fbRedFailover(i_stEntry := TC_EVENTS.PmsSystem.RedFailover);
_fbRedFailback(i_stEntry := TC_EVENTS.PmsSystem.RedFailback);
_fbRedYield(i_stEntry := TC_EVENTS.PmsSystem.RedYield);
_fbRedResume(i_stEntry := TC_EVENTS.PmsSystem.RedResume);
_fbRedSyncApplied(i_stEntry := TC_EVENTS.PmsSystem.RedSyncApplied);
_fbModeForced(i_stEntry := TC_EVENTS.PmsSeq.ModeForced);
_fbCmChange(i_stEntry := TC_EVENTS.PmsSeq.CtrlModeChange);		// [7번 수정 2026-11-09]
_fbCmRefused(i_stEntry := TC_EVENTS.PmsSeq.CtrlModeRefused);
_fbCmExit(i_stEntry := TC_EVENTS.PmsSeq.CtrlModeExit);

(* ===== 기록 구간: 아래 순서대로 한 번씩 (순서는 예전 본문과 같음) ===== *)
A_LogSystem();		// 시스템: 설정 오류·PMS 시작·운영 설정
A_LogRedundancy();	// 이중화: 절체·복귀·끊김·동기화
A_LogProtection();		// 보호 알람
A_LogDeviceFail();		// 명령 실패·장비 쓰기 실패
A_LogSource();		// 지령원 요청·끊김, 코어 상태 요청
A_LogRefused();		// 무시한 지령·기동 조건 대기·지령값 이상·배터리 요청 거부
A_LogOutput();		// 출력 제한, 자세한 기록

(* ===== 제어 모드 (메시지): 스스로 끝남 → 요청 거부 → 켜진 모드 바뀜 (전환 중 0을 내는 동안은 기다렸다가 끝난 뒤 한 번) [7번 수정 2026-11-09: 추가] ===== *)
IF iq_fbCtrlMode.q_bExitedNow THEN
	_asArg[1] := STRING_TO_WSTRING(iq_fbCtrlMode.ModuleName);
	_asArg[2] := iq_fbCtrlMode.M_SlotName(i_nSlot := iq_fbCtrlMode.q_nExitSlot);
	_asArg[3] := iq_fbCtrlMode.M_ModeReasonText(i_nSlot := iq_fbCtrlMode.q_nExitSlot, i_nReason := iq_fbCtrlMode.q_nExitReason);
	IF iq_fbCtrlMode.q_eStep = E_CtrlModeStep.Leaving THEN
		_asArg[4] := iq_fbCtrlMode.M_SlotName(i_nSlot := iq_fbCtrlMode.q_nTarget);	// 대체 모드로 가는 중
	ELSE
		_asArg[4] := iq_fbCtrlMode.M_SlotName(i_nSlot := iq_fbCtrlMode.q_nActive);
	END_IF
	_fbCmExit.M_SendEvent(4, _asArg);
END_IF
IF iq_fbCtrlMode.q_bRefusedNow THEN
	_asArg[1] := STRING_TO_WSTRING(iq_fbCtrlMode.ModuleName);
	_asArg[2] := iq_fbCtrlMode.M_SlotName(i_nSlot := iq_fbCtrlMode.q_nRefuseSlot);
	_asArg[3] := iq_fbCtrlMode.M_RefuseText();
	_fbCmRefused.M_SendEvent(3, _asArg);
END_IF
IF iq_fbCtrlMode.q_eStep <> E_CtrlModeStep.Leaving AND iq_fbCtrlMode.q_nActive <> _nCmLogged THEN
	_asArg[1] := STRING_TO_WSTRING(iq_fbCtrlMode.ModuleName);
	_asArg[2] := iq_fbCtrlMode.M_SlotName(i_nSlot := _nCmLogged);
	_asArg[3] := iq_fbCtrlMode.M_SlotName(i_nSlot := iq_fbCtrlMode.q_nActive);
	_fbCmChange.M_SendEvent(3, _asArg);
	_nCmLogged := iq_fbCtrlMode.q_nActive;
END_IF

(* ===== MQTT 브로커 끊김 (알람) [9번 수정 2026-11-09: 추가] ===== *)
IF _fbBrokerLost.q_bRaised <> i_bBrokerLost THEN
	_asArg[1] := i_sBrokerName;
	_asArg[2] := i_sBrokerDelay;
END_IF
_fbBrokerLost(i_stEntry := TC_EVENTS.PmsOutput.BrokerLost, i_bActive := i_bBrokerLost, i_nArgs := 2, i_asArg := _asArg);

_bInit := TRUE;

METHOD PRIVATE M_FillProtArgs		// 보호 알람 인자: 모듈 이름, 모듈 ID, 대상, PCS 조치, 배터리 조치
VAR_INPUT
	i_nModule	: UINT;
	i_sTarget	: WSTRING(31);
	i_stCfg		: ST_ProtCfg;
END_VAR
VAR_IN_OUT
	iq_asArg	: ARRAY[1..6] OF WSTRING(63);
END_VAR
iq_asArg[1] := M_ModuleName(i_nModule);
iq_asArg[2] := TO_WSTRING(i_nModule);
iq_asArg[3] := i_sTarget;
iq_asArg[4] := F_TxtPcsAction(i_stCfg.ePcsAction);
iq_asArg[5] := F_TxtBatAction(i_stCfg.eBatAction);
END_METHOD

METHOD PRIVATE M_IsLoggedStage : BOOL		// 로그에 남기는 단계 (요청 없음·운전 아님·램프는 정상 동작이라 안 남김)
VAR_INPUT
	i_eStage	: E_DiagStage;
END_VAR
M_IsLoggedStage := i_eStage = E_DiagStage.PccLimit OR i_eStage = E_DiagStage.DeviceLimit OR i_eStage = E_DiagStage.UnitLimit;
END_METHOD

METHOD PRIVATE M_ModuleName : WSTRING(63)	// 모듈 ID → 이름 (등록된 모듈 목록에서 찾음)
VAR_INPUT
	i_nModule	: UINT;
END_VAR
VAR
	i	: UINT;
END_VAR
M_ModuleName := WCONCAT("모듈 ", TO_WSTRING(i_nModule));
IF i_nModule = 0 THEN
	M_ModuleName := "코어";
	RETURN;
END_IF
FOR i := 1 TO GVL_PARAM.MODULE_MAX DO
	IF _aipModule[i] <> 0 AND_THEN _aipModule[i].ModuleId = i_nModule THEN
		M_ModuleName := STRING_TO_WSTRING(_aipModule[i].ModuleName);
		RETURN;
	END_IF
END_FOR
END_METHOD

METHOD PRIVATE M_ProtEventBySeverity : TcEventEntry		// 보호 이벤트 + 조치에 맞는 심각도
VAR_INPUT
	i_stCfg		: ST_ProtCfg;
END_VAR
M_ProtEventBySeverity := TC_EVENTS.PmsProt.ProtActive;
IF i_stCfg.ePcsAction = E_PcsAction.EStop OR i_stCfg.eBatAction = E_BatAction.EStop THEN
	M_ProtEventBySeverity.eSeverity := TcEventSeverity.Critical;
ELSIF i_stCfg.ePcsAction = E_PcsAction.Stop OR i_stCfg.eBatAction = E_BatAction.Stop THEN
	M_ProtEventBySeverity.eSeverity := TcEventSeverity.Error;
ELSE
	M_ProtEventBySeverity.eSeverity := TcEventSeverity.Warning;
END_IF
END_METHOD

METHOD PRIVATE M_ReasonText : WSTRING(63)	// "모듈 이름: 이유 문구" (모듈이 M_ReasonText로 직접 돌려준 문구. 모듈 0 = 코어 이유)
VAR_INPUT
	i_nModule	: UINT;
	i_nReason	: UINT;
END_VAR
VAR
	i	: UINT;
END_VAR
IF i_nModule = 0 THEN
	M_ReasonText := F_TxtCoreReason(i_nReason);
	RETURN;
END_IF
M_ReasonText := M_ModuleName(i_nModule);
FOR i := 1 TO GVL_PARAM.MODULE_MAX DO
	IF _aipModule[i] <> 0 AND_THEN _aipModule[i].ModuleId = i_nModule THEN
		M_ReasonText := WCONCAT(M_ReasonText, WCONCAT(": ", _aipModule[i].M_ReasonText(i_nReason)));
		RETURN;
	END_IF
END_FOR
END_METHOD

METHOD PRIVATE M_RuleTarget : WSTRING(31)		// 보호 대상 문구 (범위 + 대상 번호)
VAR_INPUT
	i_eScope	: E_ProtScope;
	i_nTarget	: UINT;
END_VAR
CASE i_eScope OF
	E_ProtScope.Unit:		M_RuleTarget := F_TxtNum("유닛 ", i_nTarget);
	E_ProtScope.Bms:		M_RuleTarget := F_TxtNum("BMS ", i_nTarget);
	E_ProtScope.BatGroup:	M_RuleTarget := F_TxtNum("배터리 그룹 ", i_nTarget);
	E_ProtScope.Group:		M_RuleTarget := F_TxtNum("그룹 ", i_nTarget);
ELSE
	M_RuleTarget := "사이트";
END_CASE
END_METHOD

METHOD PRIVATE M_SameLimitReason : BOOL		// 기록 기준(단계·모듈·이유)이 같은가. 값은 안 봄
VAR_INPUT
	i_stDiagA		: ST_OutputDiag;
	i_stDiagB		: ST_OutputDiag;
END_VAR
M_SameLimitReason := i_stDiagA.eStage = i_stDiagB.eStage AND i_stDiagA.nModule = i_stDiagB.nModule AND i_stDiagA.nReason = i_stDiagB.nReason
					AND i_stDiagA.eUnitBy = i_stDiagB.eUnitBy;
END_METHOD

ACTION A_LogSystem:
// 시스템: 설정 오류·PMS 시작·운영 설정
(* ===== 0-1) 설정 오류: 문구(메시지, 내용이 바뀔 때만, 처음 스캔 포함, 최대 10건), 장비 제어 중지(알람) ===== *)
_bCfgChanged := NOT _bCfgStarted OR i_nConfigErrors <> _nCfgLogged;
FOR _i := 1 TO MIN(i_nConfigErrors, 10) DO
	IF iq_asConfigErrors[_i] <> _asCfgLogged[_i] THEN
		_bCfgChanged := TRUE;
	END_IF
END_FOR
IF _bCfgChanged THEN
	FOR _i := 1 TO MIN(i_nConfigErrors, 10) DO
		_asArg[1] := iq_asConfigErrors[_i];
		_fbConfigError.M_SendEvent(1, _asArg);
		_asCfgLogged[_i] := iq_asConfigErrors[_i];
	END_FOR
	_nCfgLogged := i_nConfigErrors;
END_IF
_bCfgStarted := TRUE;
IF _fbControlBlocked.q_bRaised <> (i_nConfigErrors > 0) THEN
	_asArg[1] := TO_WSTRING(i_nConfigErrors);
END_IF
_fbControlBlocked(i_stEntry := TC_EVENTS.PmsSystem.ControlBlocked, i_bActive := i_nConfigErrors > 0, i_nArgs := 1, i_asArg := _asArg);
_fbSetRejected(i_stEntry := TC_EVENTS.PmsSystem.SettingRejected);

(* ===== 0-0) PMS 시작: 직전 동작 시각과 꺼져 있던 시간 (FB_AliveRecorder가 알려 줌) ===== *)
IF i_bPmsStart THEN
	_asArg[1] := i_sStartLastAlive;
	_asArg[2] := i_sStartOffTime;
	_fbPmsStart.M_SendEvent(2, _asArg);
END_IF

(* ===== 0) 운영 설정: 잘못된 값 되돌림(메시지), 바뀜(메시지, 저장할 때 1회), 저장 실패(알람) ===== *)
IF i_bSetRejected THEN
	_asArg[1] := i_sSetRejected;
	_fbSetRejected.M_SendEvent(1, _asArg);
END_IF
IF i_bSetChanged THEN
	_asArg[1] := i_sSetChanged;
	_fbSetChanged.M_SendEvent(1, _asArg);
END_IF
IF _fbPersistFail.q_bRaised <> i_bPersistError THEN
	_asArg[1] := TO_WSTRING(i_nPersistErrorId);
END_IF
_fbPersistFail(i_stEntry := TC_EVENTS.PmsSystem.PersistSaveFail, i_bActive := i_bPersistError, i_nArgs := 1, i_asArg := _asArg);
END_ACTION

ACTION A_LogRedundancy:
// 이중화: Active가 바뀜(메시지), 상대 끊김·통신 한쪽 고장·동기화 끊김·설정 오류(알람), 설정 맞춤(메시지)
IF NOT _bRedInit THEN
	_nRedSwitchLast		:= i_nSwitchCount;		// 시작 전에 있었던 일은 기록하지 않음
	_nRedResumeLast		:= i_nResumeCount;
	_nRedAppliedLast	:= i_nSyncApplied;
	_bRedInit			:= TRUE;
END_IF

(* 멈췄다 이어짐: 상태가 Init으로 돌아가면서 Active 횟수도 오르는데 이유는 옛 값 그대로라, 이 직후 절체 기록은 건너뜀 *)
IF i_nResumeCount <> _nRedResumeLast THEN
	_nRedResumeLast := i_nResumeCount;
	_asArg[1] := TO_WSTRING(i_nResumeCount);
	_fbRedResume.M_SendEvent(1, _asArg);
	_bRedQuiet := TRUE;
END_IF
_tonRedQuiet(IN := _bRedQuiet, PT := T#500MS);
IF _tonRedQuiet.Q THEN
	_bRedQuiet := FALSE;
END_IF

(* Active가 바뀜: 횟수가 바뀐 다음 스캔에 이유를 읽음 (횟수와 이유가 다른 태스크에서 따로 쓰여서 한 스캔 기다림) *)
IF _bRedSwitchPending THEN
	_bRedSwitchPending := FALSE;
	IF NOT _bRedQuiet THEN
		IF i_eRedRole = E_RedRole.Primary THEN
			_asArg[1] := "Primary";
		ELSE
			_asArg[1] := "Secondary";
		END_IF
		CASE i_eSwitch OF
		E_RedSwitch.Start:		_fbRedStart.M_SendEvent(1, _asArg);
		E_RedSwitch.PeerLost:	_fbRedFailover.M_SendEvent(1, _asArg);
		E_RedSwitch.Failback:	_fbRedFailback.M_SendEvent(1, _asArg);
		E_RedSwitch.Yield:		_fbRedYield.M_SendEvent(1, _asArg);
		END_CASE
	END_IF
END_IF
IF i_nSwitchCount <> _nRedSwitchLast THEN
	_nRedSwitchLast := i_nSwitchCount;
	_bRedSwitchPending := TRUE;
END_IF

